METHOD PRIVATE Test_UnconnectedMon2IsRefused
TcUnit.TEST(__POUNAME());
// arrange / act: Mon2 is unconnected, which the Safety Editor refuses
group_3(Run := TRUE);
fb_3(Mon1 := TRUE);
group_3(Run := TRUE);
fb_3(Mon1 := TRUE);
// assert
AssertEquals_BOOL(Expected := TRUE, Actual := fb_3.Error, Message := 'configuration error reported');
AssertEquals_BYTE(Expected := TO_BYTE(E_SafeFbState.Error), Actual := fb_3.State, Message := 'state ERROR');
AssertEquals_WORD(Expected := WORD#16#8000, Actual := fb_3.Diag, Message := 'diag bit 15 configuration refused');
AssertEquals_BOOL(Expected := TRUE, Actual := group_3.FbErr, Message := 'the group sees an FB error');
// act: ErrAck 0 -> 1 -> 0 does not clear a configuration error
group_3(Run := TRUE, ErrAck := TRUE);
fb_3(Mon1 := TRUE);
group_3(Run := TRUE, ErrAck := TRUE);
fb_3(Mon1 := TRUE);
group_3(Run := TRUE, ErrAck := FALSE);
fb_3(Mon1 := TRUE);
AssertEquals_BOOL(Expected := TRUE, Actual := fb_3.Error, Message := 'error not acknowledged');
AssertEquals_WORD(Expected := WORD#16#8000, Actual := fb_3.Diag, Message := 'diag bit 15 kept');
TEST_FINISHED_NAMED(__POUNAME());
END_METHOD

END_FUNCTION_BLOCK

// ---- FunctionBlocks/T_SafeEdm.TcPOU
// Model of the TwinSAFE FB EDM (external device monitor):
// Mon2 must take the opposite value to Mon1 within the configured switch-on / switch-off time.
// The Safety Editor refuses an EDM with Mon1 or Mon2 unconnected: the model then reports Error with
// diagnostic bit 15 instead of running (see T_SafeFunctionBlockBase).
{attribute 'reflection'}
FUNCTION_BLOCK T_SafeEdm EXTENDS T_SafeFunctionBlockBase
VAR_INPUT
    Mon1 : BOOL;
    Mon2 : BOOL;
    Parameters : ST_SafeEdmParameters;
END_VAR
VAR
    {attribute 'is_connected' := 'Mon1'}
    _mon1Connected : BOOL;
    {attribute 'is_connected' := 'Mon2'}
    _mon2Connected : BOOL;
    _state : E_SafeEdmState := E_SafeEdmState.Stop;
    _prevState : E_SafeEdmState;
    _timer : TON;
    _satisfied : BOOL;
END_VAR

SUPER^();
IsRunning := (_state = E_SafeEdmState.MonOn) OR (_state = E_SafeEdmState.MonOff);

// Mon1 and Mon2 must both be connected (Safety Editor: "Inport Mon1 of EDM must be connected").
METHOD PROTECTED ConfigurationOk : BOOL
IF NOT _mon1Connected THEN
    _configurationFault := 'T_SafeEdm: Inport Mon1 of EDM must be connected';
    RETURN;
ELSIF NOT _mon2Connected THEN
    _configurationFault := 'T_SafeEdm: Inport Mon2 of EDM must be connected';
    RETURN;
END_IF

ConfigurationOk := TRUE;
END_METHOD

METHOD PROTECTED Process
VAR
    monitor1 : BOOL;
    monitor2 : BOOL;
    stateBefore : E_SafeEdmState;
    passes : USINT;
END_VAR
monitor1 := F_SafeInputValue(_mon1Connected, Parameters.Mon1MakeContact, Mon1);
monitor2 := F_SafeInputValue(_mon2Connected, Parameters.Mon2MakeContact, Mon2);

IF NOT _fbRun AND _state <> E_SafeEdmState.Error AND _state <> E_SafeEdmState.Reset THEN
    _state := E_SafeEdmState.Stop;
END_IF

passes := 0;

REPEAT
    stateBefore := _state;

    CASE _state OF
        E_SafeEdmState.Stop:
            IF StateChanged() THEN
                Error := FALSE;
                Diag  := 0;
                _timer(IN := FALSE, PT := T#0S);
            END_IF

            IF _fbRun THEN
                _state := SEL(monitor1, E_SafeEdmState.MonOff, E_SafeEdmState.MonOn);
            END_IF

        E_SafeEdmState.MonOn:
            // switch-on monitoring: Mon2 must become FALSE within SwitchOnTime
            IF StateChanged() THEN
                _satisfied := FALSE;
                _timer(IN := FALSE, PT := Parameters.SwitchOnTime);
            END_IF

            IF NOT monitor2 THEN
                _satisfied := TRUE;
            END_IF

            _timer(IN := NOT _satisfied AND (Parameters.SwitchOnTime > T#0S), PT := Parameters.SwitchOnTime);

            IF _timer.Q THEN
                SetDiagBit(1);
                _state := E_SafeEdmState.Error;
            ELSIF NOT monitor1 THEN
                _state := E_SafeEdmState.MonOff;
            END_IF

        E_SafeEdmState.MonOff:
            // switch-off monitoring: Mon2 must become TRUE within SwitchOffTime
            IF StateChanged() THEN
                _satisfied := FALSE;
                _timer(IN := FALSE, PT := Parameters.SwitchOffTime);
            END_IF

            IF monitor2 THEN
                _satisfied := TRUE;
            END_IF

            _timer(IN := NOT _satisfied AND (Parameters.SwitchOffTime > T#0S), PT := Parameters.SwitchOffTime);

            IF _timer.Q THEN
                SetDiagBit(0);
                _state := E_SafeEdmState.Error;
            ELSIF monitor1 THEN
                _state := E_SafeEdmState.MonOn;
            END_IF

        E_SafeEdmState.Error:
            IF StateChanged() THEN
                Error := TRUE;
                _timer(IN := FALSE, PT := T#0S);
            END_IF

            IF _errAck THEN
                _state := E_SafeEdmState.Reset;
            END_IF

        E_SafeEdmState.Reset:
            IF StateChanged() THEN
                Error := FALSE;
                Diag  := 0;
            END_IF

            IF _errAckFallingEdge THEN
                IF NOT _fbRun THEN
                    _state := E_SafeEdmState.Stop;
                ELSE
                    _state := SEL(monitor1, E_SafeEdmState.MonOff, E_SafeEdmState.MonOn);
                END_IF
            END_IF
    END_CASE

    passes := passes + 1;
UNTIL (stateBefore = _state) OR (passes >= 3)
END_REPEAT

State := TO_BYTE(_state);
END_METHOD

METHOD PRIVATE StateChanged : BOOL
IF _prevState = _state THEN
    RETURN;
END_IF

_prevState   := _state;
StateChanged := TRUE;
END_METHOD

END_FUNCTION_BLOCK

// ---- Tests/T_SafeEStop_Tests.TcPOU
FUNCTION_BLOCK T_SafeEStop_Tests EXTENDS TcUnit.FB_TestSuite
VAR
    // Test_OutputsOffWhenStopped
    group_1 : T_SafeGroup;
    fb_1 : T_SafeEStop(group := group_1);
    // Test_StartupRequiresRestartSequence
    group_2 : T_SafeGroup;
    fb_2 : T_SafeEStop(group := group_2);
    // Test_EStopRequestSwitchesOutputsOffAndBlocksRestart
    group_3 : T_SafeGroup;
    fb_3 : T_SafeEStop(group := group_3);
    // Test_MakeContactInputRequestsSafeStateOnOne
    group_4 : T_SafeGroup;
    fb_4 : T_SafeEStop(group := group_4) := (Parameters := (EStopIn1MakeContact := TRUE));
    // Test_EdmErrorAtRestartAndAcknowledge
    group_5 : T_SafeGroup;
    fb_5 : T_SafeEStop(group := group_5);
    // Test_RestartHeldBeforeEStopGivesEdmError
    group_6 : T_SafeGroup;
    fb_6 : T_SafeEStop(group := group_6);
    // Test_DelayedOutput
    group_7 : T_SafeGroup;
    fb_7 : T_SafeEStop(group := group_7) := (Parameters := (DelayTime := T#150MS));
    state_7 : INT := 10;
    waitTimer_7 : TON;
    // Test_DiscrepancyErrorNeedsSafeInputsBeforeAck
    group_8 : T_SafeGroup;
    fb_8 : T_SafeEStop(group := group_8) := (Parameters := (DiscrepancyTime1 := T#100MS));
    state_8 : INT := 10;
    waitTimer_8 : TON;
    // Test_ResetTimeOverSixtySecondsIsRefused
    group_9 : T_SafeGroup;
    fb_9 : T_SafeEStop(group := group_9) := (Parameters := (Edm2ResetTime := T#60010MS));
END_VAR

Test_OutputsOffWhenStopped();
Test_StartupRequiresRestartSequence();
Test_EStopRequestSwitchesOutputsOffAndBlocksRestart();
Test_MakeContactInputRequestsSafeStateOnOne();
Test_EdmErrorAtRestartAndAcknowledge();
Test_RestartHeldBeforeEStopGivesEdmError();
Test_DelayedOutput();
Test_DiscrepancyErrorNeedsSafeInputsBeforeAck();
Test_ResetTimeOverSixtySecondsIsRefused();

METHOD PRIVATE Test_DelayedOutput
TcUnit.TEST(__POUNAME());
waitTimer_7();

CASE state_7 OF
    10:
        // arrange: running
        group_7(Run := TRUE);
        fb_7(Restart := FALSE, EStopIn1 := TRUE);
        group_7(Run := TRUE);
        fb_7(Restart := TRUE, EStopIn1 := TRUE);
        group_7(Run := TRUE);
        fb_7(Restart := FALSE, EStopIn1 := TRUE);
        // act
        group_7(Run := TRUE);
        fb_7(Restart := FALSE, EStopIn1 := FALSE);
        // assert
        AssertEquals_BOOL(Expected := FALSE, Actual := fb_7.EStopOut, Message := 'EStopOut off immediately');
        AssertEquals_BOOL(Expected := TRUE, Actual := fb_7.EStopDelOut, Message := 'EStopDelOut still on');
        AssertEquals_BYTE(Expected := TO_BYTE(E_SafeFbState.DelayOut), Actual := fb_7.State, Message := 'state DELAYOUT');
        state_7 := 20;
        waitTimer_7(IN := TRUE, PT := T#300MS);
    20:
        group_7(Run := TRUE);
        fb_7(Restart := FALSE, EStopIn1 := FALSE);

        IF NOT waitTimer_7.Q THEN
            RETURN;
        END_IF

        waitTimer_7(IN := FALSE);
        // assert
        AssertEquals_BOOL(Expected := FALSE, Actual := fb_7.EStopDelOut, Message := 'EStopDelOut off after the delay');
        AssertEquals_BYTE(Expected := TO_BYTE(E_SafeFbState.Safe), Actual := fb_7.State, Message := 'state SAFE');
        TEST_FINISHED_NAMED(__POUNAME());
        state_7 := 10;
END_CASE
END_METHOD

METHOD PRIVATE Test_DiscrepancyErrorNeedsSafeInputsBeforeAck
TcUnit.TEST(__POUNAME());
waitTimer_8();

CASE state_8 OF
    10:
        // arrange: running
        group_8(Run := TRUE, ErrAck := FALSE);
        fb_8(Restart := FALSE, EStopIn1 := TRUE, EStopIn2 := TRUE);
        group_8(Run := TRUE, ErrAck := FALSE);
        fb_8(Restart := TRUE, EStopIn1 := TRUE, EStopIn2 := TRUE);
        group_8(Run := TRUE, ErrAck := FALSE);
        fb_8(Restart := FALSE, EStopIn1 := TRUE, EStopIn2 := TRUE);
        state_8 := 20;
        waitTimer_8(IN := TRUE, PT := T#250MS);
    20:
        // act: only one channel opens
        group_8(Run := TRUE, ErrAck := FALSE);
        fb_8(Restart := FALSE, EStopIn1 := FALSE, EStopIn2 := TRUE);

        IF NOT waitTimer_8.Q THEN
            RETURN;
        END_IF

        waitTimer_8(IN := FALSE);
        // assert
        AssertEquals_BOOL(Expected := TRUE, Actual := fb_8.Error, Message := 'discrepancy error');
        AssertEquals_WORD(Expected := WORD#16#0101, Actual := fb_8.Diag, Message := 'diag bits 0 and 8');
        // act: acknowledge while channel 2 is still closed
        group_8(Run := TRUE, ErrAck := TRUE);
        fb_8(Restart := FALSE, EStopIn1 := FALSE, EStopIn2 := TRUE);
        AssertEquals_BYTE(Expected := TO_BYTE(E_SafeFbState.Error), Actual := fb_8.State, Message := 'ack refused until both channels safe');
        group_8(Run := TRUE, ErrAck := TRUE);
        fb_8(Restart := FALSE, EStopIn1 := FALSE, EStopIn2 := FALSE);
        AssertEquals_BYTE(Expected := TO_BYTE(E_SafeFbState.Reset), Actual := fb_8.State, Message := 'RESET once both channels were safe');
        TEST_FINISHED_NAMED(__POUNAME());
        state_8 := 10;
END_CASE
END_METHOD

METHOD PRIVATE Test_EdmErrorAtRestartAndAcknowledge
TcUnit.TEST(__POUNAME());
// arrange: EDM1 connected but contactor not released
group_5(Run := TRUE, ErrAck := FALSE);
fb_5(Restart := FALSE, EDM1 := FALSE, EStopIn1 := TRUE);
// act: restart
group_5(Run := TRUE, ErrAck := FALSE);
fb_5(Restart := TRUE, EDM1 := FALSE, EStopIn1 := TRUE);
// assert
AssertEquals_BOOL(Expected := TRUE, Actual := fb_5.Error, Message := 'EDM error when feedback missing at restart');
AssertEquals_BYTE(Expected := TO_BYTE(E_SafeFbState.Error), Actual := fb_5.State, Message := 'state ERROR');
AssertEquals_WORD(Expected := WORD#16, Actual := fb_5.Diag, Message := 'diag bit 4 EDM1');
// act: the group_5 sees the error and leaves RUN; the FB error is held
group_5(Run := TRUE, ErrAck := FALSE);
fb_5(Restart := FALSE, EDM1 := FALSE, EStopIn1 := TRUE);
AssertEquals_BYTE(Expected := TO_BYTE(E_SafeGroupState.Error), Actual := group_5.State, Message := 'group ERROR');
AssertEquals_BYTE(Expected := TO_BYTE(E_SafeFbState.Error), Actual := fb_5.State, Message := 'error is held while the group is in ERROR');
// act: ErrAck 0 -> 1 (two cycles, the group_5 needs the second to reach RESET) -> 0
group_5(Run := TRUE, ErrAck := TRUE);
fb_5(Restart := FALSE, EDM1 := FALSE, EStopIn1 := TRUE);
AssertEquals_BYTE(Expected := TO_BYTE(E_SafeFbState.Reset), Actual := fb_5.State, Message := 'state RESET while ErrAck is 1');
AssertEquals_BOOL(Expected := FALSE, Actual := fb_5.Error, Message := 'Error output off in RESET');
group_5(Run := TRUE, ErrAck := TRUE);
fb_5(Restart := FALSE, EDM1 := FALSE, EStopIn1 := TRUE);
AssertEquals_BYTE(Expected := TO_BYTE(E_SafeGroupState.Reset), Actual := group_5.State, Message := 'group RESET');
group_5(Run := TRUE, ErrAck := FALSE);
fb_5(Restart := FALSE, EDM1 := FALSE, EStopIn1 := TRUE);
AssertEquals_BYTE(Expected := TO_BYTE(E_SafeGroupState.Run), Actual := group_5.State, Message := 'group RUN after ErrAck falling edge');
AssertEquals_BYTE(Expected := TO_BYTE(E_SafeFbState.Safe), Actual := fb_5.State, Message := 'state SAFE after ErrAck falling edge');
TEST_FINISHED_NAMED(__POUNAME());
END_METHOD

METHOD PRIVATE Test_EStopRequestSwitchesOutputsOffAndBlocksRestart
TcUnit.TEST(__POUNAME());
// arrange: running
group_3(Run := TRUE);
fb_3(Restart := FALSE, EStopIn1 := TRUE, EStopIn2 := TRUE);
group_3(Run := TRUE);
fb_3(Restart := TRUE, EStopIn1 := TRUE, EStopIn2 := TRUE);
group_3(Run := TRUE);
fb_3(Restart := FALSE, EStopIn1 := TRUE, EStopIn2 := TRUE);
// act: press the e-stop
group_3(Run := TRUE);
fb_3(Restart := FALSE, EStopIn1 := FALSE, EStopIn2 := FALSE);
// assert
AssertEquals_BOOL(Expected := FALSE, Actual := fb_3.EStopOut, Message := 'EStopOut off');
AssertEquals_BOOL(Expected := FALSE, Actual := fb_3.EStopDelOut, Message := 'EStopDelOut off without delay time');
AssertEquals_BYTE(Expected := TO_BYTE(E_SafeFbState.Safe), Actual := fb_3.State, Message := 'state SAFE');
// act: restart while still pressed
group_3(Run := TRUE);
fb_3(Restart := TRUE, EStopIn1 := FALSE, EStopIn2 := FALSE);
group_3(Run := TRUE);
fb_3(Restart := FALSE, EStopIn1 := FALSE, EStopIn2 := FALSE);
AssertEquals_BOOL(Expected := FALSE, Actual := fb_3.EStopOut, Message := 'restart ignored while the e-stop is pressed');
TEST_FINISHED_NAMED(__POUNAME());
END_METHOD

METHOD PRIVATE Test_MakeContactInputRequestsSafeStateOnOne
TcUnit.TEST(__POUNAME());
// arrange: single channel make contact, released (0), restarted
group_4(Run := TRUE);
fb_4(Restart := FALSE, EStopIn1 := FALSE);
group_4(Run := TRUE);
fb_4(Restart := TRUE, EStopIn1 := FALSE);
group_4(Run := TRUE);
fb_4(Restart := FALSE, EStopIn1 := FALSE);
AssertEquals_BYTE(Expected := TO_BYTE(E_SafeFbState.Run), Actual := fb_4.State, Message := 'running with make contact released');
// act
group_4(Run := TRUE);
fb_4(Restart := FALSE, EStopIn1 := TRUE);
// assert
AssertEquals_BYTE(Expected := TO_BYTE(E_SafeFbState.Safe), Actual := fb_4.State, Message := 'make contact at 1 requests the safe state');
TEST_FINISHED_NAMED(__POUNAME());
END_METHOD

METHOD PRIVATE Test_OutputsOffWhenStopped
TcUnit.TEST(__POUNAME());
// act
group_1(Run := FALSE);
fb_1(EStopIn1 := TRUE);
// assert
AssertEquals_BOOL(Expected := FALSE, Actual := fb_1.EStopOut, Message := 'no output while the group is stopped');
AssertEquals_BYTE(Expected := TO_BYTE(E_SafeFbState.Stop), Actual := fb_1.State, Message := 'state STOP');
TEST_FINISHED_NAMED(__POUNAME());
END_METHOD

METHOD PRIVATE Test_RestartHeldBeforeEStopGivesEdmError
TcUnit.TEST(__POUNAME());
// arrange: running with EDM feedback (contactors pulled in -> EDM1 = 0)
group_6(Run := TRUE);
fb_6(Restart := FALSE, EDM1 := TRUE, EStopIn1 := TRUE);
group_6(Run := TRUE);
fb_6(Restart := TRUE, EDM1 := TRUE, EStopIn1 := TRUE);
group_6(Run := TRUE);
fb_6(Restart := FALSE, EDM1 := TRUE, EStopIn1 := TRUE);
group_6(Run := TRUE);
fb_6(Restart := FALSE, EDM1 := FALSE, EStopIn1 := TRUE);
// act: restart held, then e-stop pressed before the contactors drop out
group_6(Run := TRUE);
fb_6(Restart := TRUE, EDM1 := FALSE, EStopIn1 := FALSE);
// assert
AssertEquals_BOOL(Expected := TRUE, Actual := fb_6.Error, Message := 'immediate EDM check with restart held (sample 3)');
TEST_FINISHED_NAMED(__POUNAME());
END_METHOD

METHOD PRIVATE Test_StartupRequiresRestartSequence
TcUnit.TEST(__POUNAME());
// act: two channel e-stop released, no restart yet
group_2(Run := TRUE);
fb_2(Restart := FALSE, EStopIn1 := TRUE, EStopIn2 := TRUE);
group_2(Run := TRUE);
fb_2(Restart := FALSE, EStopIn1 := TRUE, EStopIn2 := TRUE);
// assert
AssertEquals_BOOL(Expected := FALSE, Actual := fb_2.EStopOut, Message := 'no output before restart');
AssertEquals_BYTE(Expected := TO_BYTE(E_SafeFbState.Safe), Actual := fb_2.State, Message := 'state SAFE waiting for restart');
group_2(Run := TRUE);
fb_2(Restart := TRUE, EStopIn1 := TRUE, EStopIn2 := TRUE);
AssertEquals_BYTE(Expected := TO_BYTE(E_SafeFbState.Start), Actual := fb_2.State, Message := 'state START while restart held');
AssertEquals_BOOL(Expected := FALSE, Actual := fb_2.EStopOut, Message := 'no output while restart held');
group_2(Run := TRUE);
fb_2(Restart := FALSE, EStopIn1 := TRUE, EStopIn2 := TRUE);
AssertEquals_BYTE(Expected := TO_BYTE(E_SafeFbState.Run), Actual := fb_2.State, Message := 'state RUN after falling edge');
AssertEquals_BOOL(Expected := TRUE, Actual := fb_2.EStopOut, Message := 'EStopOut on');
AssertEquals_BOOL(Expected := TRUE, Actual := fb_2.EStopDelOut, Message := 'EStopDelOut on');
TEST_FINISHED_NAMED(__POUNAME());
END_METHOD

METHOD PRIVATE Test_ResetTimeOverSixtySecondsIsRefused
TcUnit.TEST(__POUNAME());
// arrange / act: Edm2ResetTime is 60010 ms, which the Safety Editor refuses
group_9(Run := TRUE);
fb_9(EDM2 := TRUE, EStopIn1 := TRUE);
group_9(Run := TRUE);
fb_9(EDM2 := TRUE, EStopIn1 := TRUE);
// assert
AssertEquals_BOOL(Expected := TRUE, Actual := fb_9.Error, Message := 'configuration error reported');
AssertEquals_BYTE(Expected := TO_BYTE(E_SafeFbState.Error), Actual := fb_9.State, Message := 'state ERROR');
AssertEquals_WORD(Expected := WORD#16#8000, Actual := fb_9.Diag, Message := 'diag bit 15 configuration refused');
AssertEquals_BOOL(Expected := FALSE, Actual := fb_9.EStopOut, Message := 'EStopOut stays at its safe value');
AssertEquals_BOOL(Expected := TRUE, Actual := group_9.FbErr, Message := 'the group sees an FB error');
// act: ErrAck 0 -> 1 -> 0 does not clear a configuration error
group_9(Run := TRUE, ErrAck := TRUE);
fb_9(EDM2 := TRUE, EStopIn1 := TRUE);
group_9(Run := TRUE, ErrAck := TRUE);
fb_9(EDM2 := TRUE, EStopIn1 := TRUE);
group_9(Run := TRUE, ErrAck := FALSE);
fb_9(EDM2 := TRUE, EStopIn1 := TRUE);
AssertEquals_BOOL(Expected := TRUE, Actual := fb_9.Error, Message := 'error not acknowledged');
AssertEquals_WORD(Expected := WORD#16#8000, Actual := fb_9.Diag, Message := 'diag bit 15 kept');
TEST_FINISHED_NAMED(__POUNAME());
END_METHOD

END_FUNCTION_BLOCK

// ---- FunctionBlocks/T_SafeEStop.TcPOU
// Model of the TwinSAFE FB ESTOP.
// Up to eight emergency stop inputs in four pairs, immediate and delayed outputs,
// two feedback loops (EDM) and a manual restart requiring a 0 -> 1 -> 0 sequence on Restart.
// Ports are active when connected.
// The Safety Editor refuses an EDM reset time that is not 0 ms, a multiple of 10 ms and at most 60000 ms:
// the model then reports Error with diagnostic bit 15 instead of running (see T_SafeFunctionBlockBase).
{attribute 'reflection'}
FUNCTION_BLOCK T_SafeEStop EXTENDS T_SafeFunctionBlockBase
VAR_INPUT
    Restart : BOOL; // may be a standard PLC signal
    EDM1 : BOOL; // feedback loop of EStopOut (may be a standard PLC signal)
    EDM2 : BOOL; // feedback loop of EStopDelOut (may be a standard PLC signal)
    EStopIn1 : BOOL;
    EStopIn2 : BOOL;
    EStopIn3 : BOOL;
    EStopIn4 : BOOL;
    EStopIn5 : BOOL;
    EStopIn6 : BOOL;
    EStopIn7 : BOOL;
    EStopIn8 : BOOL;
    Parameters : ST_SafeEStopParameters;
END_VAR
VAR_OUTPUT
    EStopOut : BOOL; // switches off immediately
    EStopDelOut : BOOL; // switches off after DelayTime
END_VAR
VAR
    {attribute 'is_connected' := 'Restart'}
    _restartConnected : BOOL;
    {attribute 'is_connected' := 'EDM1'}
    _eDM1Connected : BOOL;
    {attribute 'is_connected' := 'EDM2'}
    _eDM2Connected : BOOL;
    {attribute 'is_connected' := 'EStopIn1'}
    _eStopIn1Connected : BOOL;
    {attribute 'is_connected' := 'EStopIn2'}
    _eStopIn2Connected : BOOL;
    {attribute 'is_connected' := 'EStopIn3'}
    _eStopIn3Connected : BOOL;
    {attribute 'is_connected' := 'EStopIn4'}
    _eStopIn4Connected : BOOL;
    {attribute 'is_connected' := 'EStopIn5'}
    _eStopIn5Connected : BOOL;
    {attribute 'is_connected' := 'EStopIn6'}
    _eStopIn6Connected : BOOL;
    {attribute 'is_connected' := 'EStopIn7'}
    _eStopIn7Connected : BOOL;
    {attribute 'is_connected' := 'EStopIn8'}
    _eStopIn8Connected : BOOL;
    _pairs : ARRAY[1..4] OF T_SafeInputPair;
    _state : E_SafeFbState := E_SafeFbState.Stop;
    _prevState : E_SafeFbState;
    _restartPrev : BOOL;
    _delayTimer : TON;
    _edmResetTimer1 : TON;
    _edmResetTimer2 : TON;
    _edm1Dropped : BOOL;
    _edm2Dropped : BOOL;
END_VAR

SUPER^();

// The EDM reset times must be 0 ms or a multiple of 10 ms up to 60000 ms (Safety Editor: "'Reset Time' parameter ... has to be 0 ms or a multiple of 10 ms and maximal 60000 ms").
METHOD PROTECTED ConfigurationOk : BOOL
IF NOT F_SafeResetTimeOk(Parameters.Edm1ResetTime) THEN
    _configurationFault := 'T_SafeEStop: $'Reset Time$' parameter of EDM1 of ESTOP has to be 0 ms or a multiple of 10 ms and maximal 60000 ms';
    RETURN;
ELSIF NOT F_SafeResetTimeOk(Parameters.Edm2ResetTime) THEN
    _configurationFault := 'T_SafeEStop: $'Reset Time$' parameter of EDM2 of ESTOP has to be 0 ms or a multiple of 10 ms and maximal 60000 ms';
    RETURN;
END_IF

ConfigurationOk := TRUE;
END_METHOD

// Checks the EDM inputs at restart and records diagnostic bits 4/5 on failure.
METHOD PRIVATE EdmInputsOk : BOOL
EdmInputsOk := TRUE;

IF _eDM1Connected AND NOT EDM1 THEN
    SetDiagBit(4);
    EdmInputsOk := FALSE;
END_IF

IF _eDM2Connected AND NOT EDM2 THEN
    SetDiagBit(5);
    EdmInputsOk := FALSE;
END_IF
END_METHOD

// TRUE when every connected EDM input reads 1 (contactors released).
METHOD PRIVATE EdmInputsTrue : BOOL
EdmInputsTrue := (NOT _eDM1Connected OR EDM1) AND (NOT _eDM2Connected OR EDM2);
END_METHOD

// EL6910 extension: after the outputs switch on, each connected EDM input must drop to FALSE
// within its Reset Time. Returns FALSE (and sets diagnostic bits 4/5) on timeout.
METHOD PRIVATE EdmResetOk : BOOL
EdmResetOk := TRUE;

IF _eDM1Connected AND Parameters.Edm1ResetTime > T#0S THEN
    IF NOT EDM1 THEN
        _edm1Dropped := TRUE;
    END_IF

    _edmResetTimer1(IN := NOT _edm1Dropped, PT := Parameters.Edm1ResetTime);

    IF _edmResetTimer1.Q THEN
        SetDiagBit(4);
        EdmResetOk := FALSE;
    END_IF
END_IF

IF _eDM2Connected AND Parameters.Edm2ResetTime > T#0S THEN
    IF NOT EDM2 THEN
        _edm2Dropped := TRUE;
    END_IF

    _edmResetTimer2(IN := NOT _edm2Dropped, PT := Parameters.Edm2ResetTime);

    IF _edmResetTimer2.Q THEN
        SetDiagBit(5);
        EdmResetOk := FALSE;
    END_IF
END_IF
END_METHOD

PROPERTY EStopState : E_SafeFbState
GET
EStopState := _state;
END_GET
END_PROPERTY

METHOD PROTECTED Process
VAR
    i : USINT;
    acknowledge : BOOL;
    safeRequested : BOOL;
    discError : BOOL;
    restartFalling : BOOL;
    operating : BOOL;
    stateBefore : E_SafeFbState;
    passes : USINT;
END_VAR
acknowledge := (_state = E_SafeFbState.Error) AND _errAck;
_pairs[1](
    In1 := EStopIn1,
    In2 := EStopIn2,
    Active1 := _eStopIn1Connected,
    Active2 := _eStopIn2Connected,
    MakeContact1 := Parameters.EStopIn1MakeContact,
    MakeContact2 := Parameters.EStopIn2MakeContact,
    DiscrepancyTime := Parameters.DiscrepancyTime1,
    Monitor := _fbRun,
    SafeInputsAfterDiscError := TRUE, // the EL6910 always applies it to ESTOP, whatever the parameter says
    Acknowledge := acknowledge
);

_pairs[2](
    In1 := EStopIn3,
    In2 := EStopIn4,
    Active1 := _eStopIn3Connected,
    Active2 := _eStopIn4Connected,
    MakeContact1 := Parameters.EStopIn3MakeContact,
    MakeContact2 := Parameters.EStopIn4MakeContact,
    DiscrepancyTime := Parameters.DiscrepancyTime2,
    Monitor := _fbRun,
    SafeInputsAfterDiscError := TRUE, // the EL6910 always applies it to ESTOP, whatever the parameter says
    Acknowledge := acknowledge
);

_pairs[3](
    In1 := EStopIn5,
    In2 := EStopIn6,
    Active1 := _eStopIn5Connected,
    Active2 := _eStopIn6Connected,
    MakeContact1 := Parameters.EStopIn5MakeContact,
    MakeContact2 := Parameters.EStopIn6MakeContact,
    DiscrepancyTime := Parameters.DiscrepancyTime3,
    Monitor := _fbRun,
    SafeInputsAfterDiscError := TRUE, // the EL6910 always applies it to ESTOP, whatever the parameter says
    Acknowledge := acknowledge
);

_pairs[4](
    In1 := EStopIn7,
    In2 := EStopIn8,
    Active1 := _eStopIn7Connected,
    Active2 := _eStopIn8Connected,
    MakeContact1 := Parameters.EStopIn7MakeContact,
    MakeContact2 := Parameters.EStopIn8MakeContact,
    DiscrepancyTime := Parameters.DiscrepancyTime4,
    Monitor := _fbRun,
    SafeInputsAfterDiscError := TRUE, // the EL6910 always applies it to ESTOP, whatever the parameter says
    Acknowledge := acknowledge
);

FOR i := 1 TO 4 DO
    safeRequested := safeRequested OR _pairs[i].SafeStateRequested;
    discError     := discError OR _pairs[i].DiscrepancyError;
END_FOR

restartFalling := NOT Restart AND _restartPrev;
_restartPrev   := Restart;

IF NOT _fbRun AND _state <> E_SafeFbState.Error AND _state <> E_SafeFbState.Reset THEN
    _state := E_SafeFbState.Stop;
END_IF

// A discrepancy error is detected in every operating state
operating := (_state = E_SafeFbState.Safe)
                 OR (_state = E_SafeFbState.Start)
                 OR (_state = E_SafeFbState.Run)
                 OR (_state = E_SafeFbState.DelayOut);

IF discError AND operating THEN
    UpdateDiscrepancyDiag();
    _state := E_SafeFbState.Error;
END_IF

passes := 0;

REPEAT
    stateBefore := _state;

    CASE _state OF
        E_SafeFbState.Stop:
            IF StateChanged() THEN
                SetOutputsSafe();
                Error := FALSE;
                Diag  := 0;
            END_IF

            IF _fbRun THEN
                _state := E_SafeFbState.Safe;
            END_IF

        E_SafeFbState.Safe:
            IF StateChanged() THEN
                SetOutputsSafe();
            END_IF

            // A TRUE restart signal triggers the EDM check immediately (see restart behaviour sample 3)
            IF Restart THEN
                IF NOT EdmInputsOk() THEN
                    _state := E_SafeFbState.Error;
                ELSIF NOT safeRequested THEN
                    _state := E_SafeFbState.Start;
                END_IF
            END_IF

        E_SafeFbState.Start:
            IF StateChanged() THEN
                SetOutputsSafe();
            END_IF

            IF safeRequested THEN
                _state := E_SafeFbState.Safe;
            ELSIF restartFalling THEN
                IF EdmInputsOk() THEN
                    _state := E_SafeFbState.Run;
                ELSE
                    _state := E_SafeFbState.Error;
                END_IF
            END_IF

        E_SafeFbState.Run:
            IF StateChanged() THEN
                EStopOut    := TRUE;
                EStopDelOut := TRUE;
                StartEdmResetMonitoring();
            END_IF

            IF NOT EdmResetOk() THEN
                _state := E_SafeFbState.Error;
            ELSIF safeRequested THEN
                IF Parameters.DelayTime > T#0S THEN
                    _state := E_SafeFbState.DelayOut;
                ELSE
                    _state := E_SafeFbState.Safe;
                END_IF
            END_IF

        E_SafeFbState.DelayOut:
            IF StateChanged() THEN
                EStopOut    := FALSE;
                EStopDelOut := TRUE;
                _delayTimer(IN := FALSE, PT := Parameters.DelayTime);
            END_IF

            _delayTimer(IN := TRUE, PT := Parameters.DelayTime);

            IF _delayTimer.Q THEN
                _state := E_SafeFbState.Safe;
            END_IF

        E_SafeFbState.Error:
            IF StateChanged() THEN
                SetOutputsSafe();
                Error := TRUE;
            END_IF

            UpdateDiscrepancyDiag();

            IF _errAck AND NOT discError THEN
                _state := E_SafeFbState.Reset;
            END_IF

        E_SafeFbState.Reset:
            IF StateChanged() THEN
                SetOutputsSafe();
                Error := FALSE;
                Diag  := 0;
            END_IF

            IF _errAckFallingEdge THEN
                _state := SEL(_fbRun, E_SafeFbState.Stop, E_SafeFbState.Safe);
            END_IF
    END_CASE

    passes := passes + 1;
UNTIL (stateBefore = _state) OR (passes >= 3)
END_REPEAT

State := TO_BYTE(_state);
END_METHOD

METHOD PRIVATE SetOutputsSafe
EStopOut    := FALSE;
EStopDelOut := FALSE;
END_METHOD

METHOD PRIVATE StartEdmResetMonitoring
_edm1Dropped := FALSE;
_edm2Dropped := FALSE;
_edmResetTimer1(IN := FALSE, PT := Parameters.Edm1ResetTime);
_edmResetTimer2(IN := FALSE, PT := Parameters.Edm2ResetTime);
END_METHOD

METHOD PRIVATE StateChanged : BOOL
IF _prevState = _state THEN
    RETURN;
END_IF

_prevState   := _state;
StateChanged := TRUE;
END_METHOD

// Mirrors the discrepancy state of every pair into the diagnostic bits.
METHOD PRIVATE UpdateDiscrepancyDiag
VAR
    i : USINT;
END_VAR
FOR i := 1 TO 4 DO
    IF _pairs[i].DiscrepancyError THEN
        SetDiagBit(i - 1);

        IF _pairs[i].AwaitingSafeInputs THEN
            SetDiagBit(i + 7);
        ELSE
            ClearDiagBit(i + 7);
        END_IF
    END_IF
END_FOR
END_METHOD

END_FUNCTION_BLOCK

// ---- Core/F_SafeResetTimeOk.TcPOU
// TRUE when an EDM 'Reset Time' parameter is one the Safety Editor accepts: 0 ms (off) or a multiple
// of 10 ms, and at most 60000 ms. The editor reports "'Reset Time' parameter ... has to be 0 ms or a
// multiple of 10 ms and maximal 60000 ms" otherwise.
FUNCTION F_SafeResetTimeOk : BOOL
VAR_INPUT
    resetTime : TIME;
END_VAR
VAR CONSTANT
    MAX_RESET_TIME : TIME := T#60S;
END_VAR

IF resetTime > MAX_RESET_TIME THEN
    RETURN;
END_IF

F_SafeResetTimeOk := (TIME_TO_UDINT(resetTime) MOD 10 = 0);

END_FUNCTION

// ---- Tests/T_SafeMon_Tests.TcPOU
FUNCTION_BLOCK T_SafeMon_Tests EXTENDS TcUnit.FB_TestSuite
VAR
    // Test_AutomaticRestartWhenGuardClosed
    group_1 : T_SafeGroup;
    fb_1 : T_SafeMon(group := group_1);
    // Test_SecureInputBypassesGuard
    group_2 : T_SafeGroup;
    fb_2 : T_SafeMon(group := group_2);
    // Test_ManualFunctionTestRequiresGuardOpenedOnce
    group_3 : T_SafeGroup;
    fb_3 : T_SafeMon(group := group_3) := (Parameters := (ManualFunctionTest := TRUE));
    // Test_EdmFaultWithoutManualRestartStaysSafe
    group_4 : T_SafeGroup;
    fb_4 : T_SafeMon(group := group_4);
    // Test_NoMonInConnectedIsRefused
    group_5 : T_SafeGroup;
    fb_5 : T_SafeMon(group := group_5);
    // Test_ResetTimeNotMultipleOfTenIsRefused
    group_6 : T_SafeGroup;
    fb_6 : T_SafeMon(group := group_6) := (Parameters := (Edm1ResetTime := T#15MS));
END_VAR

Test_AutomaticRestartWhenGuardClosed();
Test_SecureInputBypassesGuard();
Test_ManualFunctionTestRequiresGuardOpenedOnce();
Test_EdmFaultWithoutManualRestartStaysSafe();
Test_NoMonInConnectedIsRefused();
Test_ResetTimeNotMultipleOfTenIsRefused();

METHOD PRIVATE Test_AutomaticRestartWhenGuardClosed
TcUnit.TEST(__POUNAME());
// act: Restart not connected -> automatic restart; guard open
group_1(Run := TRUE);
fb_1(MonIn1 := FALSE);
group_1(Run := TRUE);
fb_1(MonIn1 := FALSE);
// assert
AssertEquals_BOOL(Expected := FALSE, Actual := fb_1.MonOut, Message := 'output off with guard open');
group_1(Run := TRUE);
fb_1(MonIn1 := TRUE);
AssertEquals_BOOL(Expected := TRUE, Actual := fb_1.MonOut, Message := 'automatic restart with guard closed');
AssertEquals_BYTE(Expected := TO_BYTE(E_SafeMonState.Run), Actual := fb_1.State, Message := 'state RUN');
TEST_FINISHED_NAMED(__POUNAME());
END_METHOD

METHOD PRIVATE Test_EdmFaultWithoutManualRestartStaysSafe
TcUnit.TEST(__POUNAME());
// act: EDM1 connected and FALSE, no Restart connected
group_4(Run := TRUE);
fb_4(EDM1 := FALSE, MonIn1 := TRUE);
group_4(Run := TRUE);
fb_4(EDM1 := FALSE, MonIn1 := TRUE);
// assert
AssertEquals_BOOL(Expected := FALSE, Actual := fb_4.Error, Message := 'no EDM error without manual restart');
AssertEquals_BYTE(Expected := TO_BYTE(E_SafeMonState.Safe), Actual := fb_4.State, Message := 'FB remains SAFE');
TEST_FINISHED_NAMED(__POUNAME());
END_METHOD

METHOD PRIVATE Test_ManualFunctionTestRequiresGuardOpenedOnce
TcUnit.TEST(__POUNAME());
// arrange: Restart connected (manual restart), guard closed from the start
group_3(Run := TRUE);
fb_3(Restart := FALSE, MonIn1 := TRUE);
AssertEquals_BYTE(Expected := TO_BYTE(E_SafeMonState.FuncTest), Actual := fb_3.State, Message := 'state FUNCTEST after start');
// act: restart without testing the guard
group_3(Run := TRUE);
fb_3(Restart := TRUE, MonIn1 := TRUE);
group_3(Run := TRUE);
fb_3(Restart := FALSE, MonIn1 := TRUE);
AssertEquals_BOOL(Expected := FALSE, Actual := fb_3.MonOut, Message := 'restart ignored before the function test');
// act: open and close the guard, then restart
group_3(Run := TRUE);
fb_3(Restart := FALSE, MonIn1 := FALSE);
group_3(Run := TRUE);
fb_3(Restart := FALSE, MonIn1 := TRUE);
group_3(Run := TRUE);
fb_3(Restart := TRUE, MonIn1 := TRUE);
group_3(Run := TRUE);
fb_3(Restart := FALSE, MonIn1 := TRUE);
AssertEquals_BOOL(Expected := TRUE, Actual := fb_3.MonOut, Message := 'output on after function test and restart');
TEST_FINISHED_NAMED(__POUNAME());
END_METHOD

METHOD PRIVATE Test_SecureInputBypassesGuard
TcUnit.TEST(__POUNAME());
// act: guard open, bypass active
group_2(Run := TRUE);
fb_2(MonIn1 := FALSE, Secure1 := TRUE);
group_2(Run := TRUE);
fb_2(MonIn1 := FALSE, Secure1 := TRUE);
// assert
AssertEquals_BOOL(Expected := TRUE, Actual := fb_2.MonOut, Message := 'guard ignored while Secure is 1');
group_2(Run := TRUE);
fb_2(MonIn1 := FALSE, Secure1 := FALSE);
AssertEquals_BOOL(Expected := FALSE, Actual := fb_2.MonOut, Message := 'guard monitored again when Secure is 0');
TEST_FINISHED_NAMED(__POUNAME());
END_METHOD

METHOD PRIVATE Test_NoMonInConnectedIsRefused
TcUnit.TEST(__POUNAME());
// arrange / act: only the Secure pair is connected, which the Safety Editor refuses
group_5(Run := TRUE);
fb_5(Secure1 := TRUE);
group_5(Run := TRUE);
fb_5(Secure1 := TRUE);
// assert
AssertEquals_BOOL(Expected := TRUE, Actual := fb_5.Error, Message := 'configuration error reported');
AssertEquals_BYTE(Expected := TO_BYTE(E_SafeFbState.Error), Actual := fb_5.State, Message := 'state ERROR');
AssertEquals_WORD(Expected := WORD#16#8000, Actual := fb_5.Diag, Message := 'diag bit 15 configuration refused');
AssertEquals_BOOL(Expected := FALSE, Actual := fb_5.MonOut, Message := 'MonOut stays at its safe value');
AssertEquals_BOOL(Expected := TRUE, Actual := group_5.FbErr, Message := 'the group sees an FB error');
// act: ErrAck 0 -> 1 -> 0 does not clear a configuration error
group_5(Run := TRUE, ErrAck := TRUE);
fb_5(Secure1 := TRUE);
group_5(Run := TRUE, ErrAck := TRUE);
fb_5(Secure1 := TRUE);
group_5(Run := TRUE, ErrAck := FALSE);
fb_5(Secure1 := TRUE);
AssertEquals_BOOL(Expected := TRUE, Actual := fb_5.Error, Message := 'error not acknowledged');
AssertEquals_WORD(Expected := WORD#16#8000, Actual := fb_5.Diag, Message := 'diag bit 15 kept');
TEST_FINISHED_NAMED(__POUNAME());
END_METHOD

METHOD PRIVATE Test_ResetTimeNotMultipleOfTenIsRefused
TcUnit.TEST(__POUNAME());
// arrange / act: Edm1ResetTime is 15 ms, which the Safety Editor refuses
group_6(Run := TRUE);
fb_6(EDM1 := TRUE, MonIn1 := TRUE);
group_6(Run := TRUE);
fb_6(EDM1 := TRUE, MonIn1 := TRUE);
// assert
AssertEquals_BOOL(Expected := TRUE, Actual := fb_6.Error, Message := 'configuration error reported');
AssertEquals_BYTE(Expected := TO_BYTE(E_SafeFbState.Error), Actual := fb_6.State, Message := 'state ERROR');
AssertEquals_WORD(Expected := WORD#16#8000, Actual := fb_6.Diag, Message := 'diag bit 15 configuration refused');
AssertEquals_BOOL(Expected := FALSE, Actual := fb_6.MonOut, Message := 'MonOut stays at its safe value');
AssertEquals_BOOL(Expected := TRUE, Actual := group_6.FbErr, Message := 'the group sees an FB error');
// act: ErrAck 0 -> 1 -> 0 does not clear a configuration error
group_6(Run := TRUE, ErrAck := TRUE);
fb_6(EDM1 := TRUE, MonIn1 := TRUE);
group_6(Run := TRUE, ErrAck := TRUE);
fb_6(EDM1 := TRUE, MonIn1 := TRUE);
group_6(Run := TRUE, ErrAck := FALSE);
fb_6(EDM1 := TRUE, MonIn1 := TRUE);
AssertEquals_BOOL(Expected := TRUE, Actual := fb_6.Error, Message := 'error not acknowledged');
AssertEquals_WORD(Expected := WORD#16#8000, Actual := fb_6.Diag, Message := 'diag bit 15 kept');
TEST_FINISHED_NAMED(__POUNAME());
END_METHOD

END_FUNCTION_BLOCK

// ---- FunctionBlocks/T_SafeMon.TcPOU
// Model of the TwinSAFE FB MON (safety door / guard monitoring).
// Two MonIn pairs, a Secure pair that bypasses them, manual restart (when Restart is connected),
// manual function test, two EDM feedback loops and a delayed output.
// The Safety Editor refuses a MON with no MonIn port connected, or an EDM reset time that is not 0 ms,
// a multiple of 10 ms and at most 60000 ms: the model then reports Error with diagnostic bit 15
// instead of running (see T_SafeFunctionBlockBase).
{attribute 'reflection'}
FUNCTION_BLOCK T_SafeMon EXTENDS T_SafeFunctionBlockBase
VAR_INPUT
    Restart : BOOL; // connect for manual restart; may be a standard PLC signal
    EDM1 : BOOL; // feedback loop of MonOut
    EDM2 : BOOL; // feedback loop of MonDelOut
    MonIn1 : BOOL;
    MonIn2 : BOOL;
    MonIn3 : BOOL;
    MonIn4 : BOOL;
    Secure1 : BOOL; // when TRUE (after normalisation) the MonIn inputs are ignored
    Secure2 : BOOL;
    Parameters : ST_SafeMonParameters;
END_VAR
VAR_OUTPUT
    MonOut : BOOL;
    MonDelOut : BOOL;
END_VAR
VAR
    {attribute 'is_connected' := 'Restart'}
    _restartConnected : BOOL;
    {attribute 'is_connected' := 'EDM1'}
    _eDM1Connected : BOOL;
    {attribute 'is_connected' := 'EDM2'}
    _eDM2Connected : BOOL;
    {attribute 'is_connected' := 'MonIn1'}
    _monIn1Connected : BOOL;
    {attribute 'is_connected' := 'MonIn2'}
    _monIn2Connected : BOOL;
    {attribute 'is_connected' := 'MonIn3'}
    _monIn3Connected : BOOL;
    {attribute 'is_connected' := 'MonIn4'}
    _monIn4Connected : BOOL;
    {attribute 'is_connected' := 'Secure1'}
    _secure1Connected : BOOL;
    {attribute 'is_connected' := 'Secure2'}
    _secure2Connected : BOOL;
    _pairs : ARRAY[1..3] OF T_SafeInputPair; // 1: MonIn1/2, 2: MonIn3/4, 3: Secure1/2
    _state : E_SafeMonState := E_SafeMonState.Stop;
    _prevState : E_SafeMonState;
    _restartPrev : BOOL;
    _delayTimer : TON;
    _delayRunning : BOOL;
    _funcTested : ARRAY[1..2] OF BOOL;
    _edmResetTimer1 : TON;
    _edmResetTimer2 : TON;
    _edm1Dropped : BOOL;
    _edm2Dropped : BOOL;
END_VAR

SUPER^();

// At least one MonIn port must be connected and the EDM reset times must be 0 ms or a multiple of 10 ms up to 60000 ms (Safety Editor messages).
METHOD PROTECTED ConfigurationOk : BOOL
IF NOT (_monIn1Connected OR _monIn2Connected OR _monIn3Connected OR _monIn4Connected) THEN
    _configurationFault := 'T_SafeMon: MON does not have at least 1 MonIn(x) port active and connected';
    RETURN;
ELSIF NOT F_SafeResetTimeOk(Parameters.Edm1ResetTime) THEN
    _configurationFault := 'T_SafeMon: $'Reset Time$' parameter of EDM1 of MON has to be 0 ms or a multiple of 10 ms and maximal 60000 ms';
    RETURN;
ELSIF NOT F_SafeResetTimeOk(Parameters.Edm2ResetTime) THEN
    _configurationFault := 'T_SafeMon: $'Reset Time$' parameter of EDM2 of MON has to be 0 ms or a multiple of 10 ms and maximal 60000 ms';
    RETURN;
END_IF

ConfigurationOk := TRUE;
END_METHOD

// Checks the EDM inputs at restart and records diagnostic bits 4/5 on failure.
METHOD PRIVATE EdmInputsOk : BOOL
EdmInputsOk := TRUE;

IF _eDM1Connected AND NOT EDM1 THEN
    SetDiagBit(4);
    EdmInputsOk := FALSE;
END_IF

IF _eDM2Connected AND NOT EDM2 THEN
    SetDiagBit(5);
    EdmInputsOk := FALSE;
END_IF
END_METHOD

// TRUE when every connected EDM input reads 1 (contactors released).
METHOD PRIVATE EdmInputsTrue : BOOL
EdmInputsTrue := (NOT _eDM1Connected OR EDM1) AND (NOT _eDM2Connected OR EDM2);
END_METHOD

// EL6910 extension: after the outputs switch on, each connected EDM input must drop to FALSE
// within its Reset Time. Returns FALSE (and sets diagnostic bits 4/5) on timeout.
METHOD PRIVATE EdmResetOk : BOOL
EdmResetOk := TRUE;

IF _eDM1Connected AND Parameters.Edm1ResetTime > T#0S THEN
    IF NOT EDM1 THEN
        _edm1Dropped := TRUE;
    END_IF

    _edmResetTimer1(IN := NOT _edm1Dropped, PT := Parameters.Edm1ResetTime);

    IF _edmResetTimer1.Q THEN
        SetDiagBit(4);
        EdmResetOk := FALSE;
    END_IF
END_IF

IF _eDM2Connected AND Parameters.Edm2ResetTime > T#0S THEN
    IF NOT EDM2 THEN
        _edm2Dropped := TRUE;
    END_IF

    _edmResetTimer2(IN := NOT _edm2Dropped, PT := Parameters.Edm2ResetTime);

    IF _edmResetTimer2.Q THEN
        SetDiagBit(5);
        EdmResetOk := FALSE;
    END_IF
END_IF
END_METHOD

PROPERTY MonState : E_SafeMonState
GET
MonState := _state;
END_GET
END_PROPERTY

METHOD PROTECTED Process
VAR
    i : USINT;
    acknowledge : BOOL;
    monRequested : BOOL;
    bypass : BOOL;
    safeRequested : BOOL;
    discError : BOOL;
    restartFalling : BOOL;
    functionTestDue : BOOL;
    stateBefore : E_SafeMonState;
    passes : USINT;
END_VAR
acknowledge := (_state = E_SafeMonState.Error) AND _errAck;
_pairs[1](
    In1 := MonIn1,
    In2 := MonIn2,
    Active1 := _monIn1Connected,
    Active2 := _monIn2Connected,
    MakeContact1 := Parameters.MonIn1MakeContact,
    MakeContact2 := Parameters.MonIn2MakeContact,
    DiscrepancyTime := Parameters.DiscrepancyTime1,
    Monitor := _fbRun,
    SafeInputsAfterDiscError := Parameters.SafeInputsAfterDiscError,
    Acknowledge := acknowledge
);

_pairs[2](
    In1 := MonIn3,
    In2 := MonIn4,
    Active1 := _monIn3Connected,
    Active2 := _monIn4Connected,
    MakeContact1 := Parameters.MonIn3MakeContact,
    MakeContact2 := Parameters.MonIn4MakeContact,
    DiscrepancyTime := Parameters.DiscrepancyTime2,
    Monitor := _fbRun,
    SafeInputsAfterDiscError := Parameters.SafeInputsAfterDiscError,
    Acknowledge := acknowledge
);

_pairs[3](
    In1 := Secure1,
    In2 := Secure2,
    Active1 := _secure1Connected,
    Active2 := _secure2Connected,
    MakeContact1 := Parameters.Secure1MakeContact,
    MakeContact2 := Parameters.Secure2MakeContact,
    DiscrepancyTime := Parameters.SecureDiscrepancyTime,
    Monitor := _fbRun,
    SafeInputsAfterDiscError := Parameters.SafeInputsAfterDiscError,
    Acknowledge := acknowledge
);

monRequested  := _pairs[1].SafeStateRequested OR _pairs[2].SafeStateRequested;
bypass        := _pairs[3].IsActive AND _pairs[3].AllTrue;
safeRequested := monRequested AND NOT bypass;

FOR i := 1 TO 3 DO
    discError := discError OR _pairs[i].DiscrepancyError;
END_FOR

restartFalling := NOT Restart AND _restartPrev;
_restartPrev   := Restart;

IF NOT _fbRun AND _state <> E_SafeMonState.Error AND _state <> E_SafeMonState.Reset THEN
    _state := E_SafeMonState.Stop;
END_IF

// Discrepancy errors: immediate, except that a running delayed output completes its delay first
IF discError THEN
    CASE _state OF
        E_SafeMonState.Safe, E_SafeMonState.Start, E_SafeMonState.FuncTest:
            UpdateDiscrepancyDiag();
            _state := E_SafeMonState.Error;
        E_SafeMonState.Run:
            UpdateDiscrepancyDiag();

            IF Parameters.DelayTime > T#0S THEN
                _state := E_SafeMonState.ErrorDelay;
            ELSE
                _state := E_SafeMonState.Error;
            END_IF
        E_SafeMonState.DelayOut:
            UpdateDiscrepancyDiag();
            _state := E_SafeMonState.ErrorDelay;
    END_CASE
END_IF

passes := 0;

REPEAT
    stateBefore := _state;

    CASE _state OF
        E_SafeMonState.Stop:
            IF StateChanged() THEN
                SetOutputsSafe();
                Error          := FALSE;
                Diag           := 0;
                _delayRunning  := FALSE;
                _funcTested[1] := FALSE;
                _funcTested[2] := FALSE;
            END_IF

            IF _fbRun THEN
                functionTestDue := Parameters.ManualFunctionTest AND (_pairs[1].IsActive OR _pairs[2].IsActive);
                _state          := SEL(functionTestDue, E_SafeMonState.Safe, E_SafeMonState.FuncTest);
            END_IF

        E_SafeMonState.FuncTest:
            // every connected MonIn pair must request the safe state once before a restart is accepted
            IF StateChanged() THEN
                SetOutputsSafe();
            END_IF

            IF _pairs[1].SafeStateRequested THEN
                _funcTested[1] := TRUE;
            END_IF

            IF _pairs[2].SafeStateRequested THEN
                _funcTested[2] := TRUE;
            END_IF

            IF (NOT _pairs[1].IsActive OR _funcTested[1]) AND (NOT _pairs[2].IsActive OR _funcTested[2]) THEN
                _state := E_SafeMonState.Safe;
            END_IF

        E_SafeMonState.Safe:
            IF StateChanged() THEN
                SetOutputsSafe();
                _delayRunning := FALSE;
            END_IF

            IF _restartConnected THEN
                IF Restart THEN
                    IF NOT EdmInputsOk() THEN
                        _state := E_SafeMonState.Error;
                    ELSIF NOT safeRequested THEN
                        _state := E_SafeMonState.Start;
                    END_IF
                END_IF
            ELSIF NOT safeRequested AND EdmInputsTrue() THEN
                // automatic restart: an EDM fault keeps the FB in SAFE without an error
                _state := E_SafeMonState.Run;
            END_IF

        E_SafeMonState.Start:
            IF StateChanged() THEN
                SetOutputsSafe();
            END_IF

            IF safeRequested THEN
                _state := E_SafeMonState.Safe;
            ELSIF restartFalling THEN
                IF EdmInputsOk() THEN
                    _state := E_SafeMonState.Run;
                ELSE
                    _state := E_SafeMonState.Error;
                END_IF
            END_IF

        E_SafeMonState.Run:
            IF StateChanged() THEN
                MonOut    := TRUE;
                MonDelOut := TRUE;
                StartEdmResetMonitoring();
            END_IF

            IF NOT EdmResetOk() THEN
                _state := E_SafeMonState.Error;
            ELSIF safeRequested THEN
                IF Parameters.DelayTime > T#0S THEN
                    _state := E_SafeMonState.DelayOut;
                ELSE
                    _state := E_SafeMonState.Safe;
                END_IF
            END_IF

        E_SafeMonState.DelayOut:
            IF StateChanged() THEN
                MonOut    := FALSE;
                MonDelOut := TRUE;
                _delayTimer(IN := FALSE, PT := Parameters.DelayTime);
                _delayRunning := TRUE;
            END_IF

            _delayTimer(IN := TRUE, PT := Parameters.DelayTime);

            IF _delayTimer.Q THEN
                _state := E_SafeMonState.Safe;
            END_IF

        E_SafeMonState.ErrorDelay:
            IF StateChanged() THEN
                MonOut    := FALSE;
                MonDelOut := TRUE;

                IF NOT _delayRunning THEN
                    _delayTimer(IN := FALSE, PT := Parameters.DelayTime);
                    _delayRunning := TRUE;
                END_IF
            END_IF

            _delayTimer(IN := TRUE, PT := Parameters.DelayTime);

            IF _delayTimer.Q THEN
                _state := E_SafeMonState.Error;
            END_IF

        E_SafeMonState.Error:
            IF StateChanged() THEN
                SetOutputsSafe();
                Error         := TRUE;
                _delayRunning := FALSE;
            END_IF

            UpdateDiscrepancyDiag();

            IF _errAck AND NOT discError THEN
                _state := E_SafeMonState.Reset;
            END_IF

        E_SafeMonState.Reset:
            IF StateChanged() THEN
                SetOutputsSafe();
                Error := FALSE;
                Diag  := 0;
            END_IF

            IF _errAckFallingEdge THEN
                _state := SEL(_fbRun, E_SafeMonState.Stop, E_SafeMonState.Safe);
            END_IF
    END_CASE

    passes := passes + 1;
UNTIL (stateBefore = _state) OR (passes >= 3)
END_REPEAT

State := TO_BYTE(_state);
END_METHOD

METHOD PRIVATE SetOutputsSafe
MonOut    := FALSE;
MonDelOut := FALSE;
END_METHOD

METHOD PRIVATE StartEdmResetMonitoring
_edm1Dropped := FALSE;
_edm2Dropped := FALSE;
_edmResetTimer1(IN := FALSE, PT := Parameters.Edm1ResetTime);
_edmResetTimer2(IN := FALSE, PT := Parameters.Edm2ResetTime);
END_METHOD

METHOD PRIVATE StateChanged : BOOL
IF _prevState = _state THEN
    RETURN;
END_IF

_prevState   := _state;
StateChanged := TRUE;
END_METHOD

// Mirrors the discrepancy state of every pair into the diagnostic bits.
METHOD PRIVATE UpdateDiscrepancyDiag
VAR
    i : USINT;
END_VAR
FOR i := 1 TO 3 DO
    IF _pairs[i].DiscrepancyError THEN
        SetDiagBit(i - 1);

        IF _pairs[i].AwaitingSafeInputs THEN
            SetDiagBit(i + 7);
        ELSE
            ClearDiagBit(i + 7);
        END_IF
    END_IF
END_FOR
END_METHOD

END_FUNCTION_BLOCK

// ---- Tests/T_SafeTwoHand_Tests.TcPOU
FUNCTION_BLOCK T_SafeTwoHand_Tests EXTENDS TcUnit.FB_TestSuite
VAR
    // Test_BothHandsGiveOutputAndReleaseNeedsBothOff
    group_1 : T_SafeGroup;
    fb_1 : T_SafeTwoHand(group := group_1);
    // Test_SecondHandWithoutFirstGivesTwoHandError
    group_2 : T_SafeGroup;
    fb_2 : T_SafeTwoHand(group := group_2);
    // Test_HandDiscrepancyTimeout
    group_3 : T_SafeGroup;
    // SafeInputsAfterDiscError TRUE (not the default) so the error waits for both hands released (diag bit 10)
    fb_3 : T_SafeTwoHand(group := group_3) := (Parameters := (HandDiscrepancyTime := T#100MS, SafeInputsAfterDiscError := TRUE));
    state_3 : INT := 10;
    waitTimer_3 : TON;
END_VAR

Test_BothHandsGiveOutputAndReleaseNeedsBothOff();
Test_SecondHandWithoutFirstGivesTwoHandError();
Test_HandDiscrepancyTimeout();

METHOD PRIVATE Test_BothHandsGiveOutputAndReleaseNeedsBothOff
TcUnit.TEST(__POUNAME());
// arrange: single channel per hand
group_1(Run := TRUE);
fb_1(Twohand1 := FALSE, Twohand3 := FALSE);
// act
group_1(Run := TRUE);
fb_1(Twohand1 := TRUE, Twohand3 := FALSE);
AssertEquals_BYTE(Expected := TO_BYTE(E_SafeTwoHandState.OneButton), Actual := fb_1.State, Message := 'state 1BUTTON');
group_1(Run := TRUE);
fb_1(Twohand1 := TRUE, Twohand3 := TRUE);
// assert
AssertEquals_BOOL(Expected := TRUE, Actual := fb_1.TwoHandOut, Message := 'output on with both hands');
group_1(Run := TRUE);
fb_1(Twohand1 := FALSE, Twohand3 := TRUE);
AssertEquals_BOOL(Expected := FALSE, Actual := fb_1.TwoHandOut, Message := 'output off when one hand released');
AssertEquals_BYTE(Expected := TO_BYTE(E_SafeTwoHandState.Release), Actual := fb_1.State, Message := 'state RELEASE');
group_1(Run := TRUE);
fb_1(Twohand1 := TRUE, Twohand3 := TRUE);
AssertEquals_BOOL(Expected := FALSE, Actual := fb_1.TwoHandOut, Message := 'no re-trigger until both hands released');
TEST_FINISHED_NAMED(__POUNAME());
END_METHOD

METHOD PRIVATE Test_HandDiscrepancyTimeout
TcUnit.TEST(__POUNAME());
waitTimer_3();

CASE state_3 OF
    10:
        group_3(Run := TRUE);
        fb_3(Twohand1 := FALSE, Twohand3 := FALSE);
        state_3 := 20;
        waitTimer_3(IN := TRUE, PT := T#250MS);
    20:
        // act: only one hand for longer than the discrepancy time
        group_3(Run := TRUE);
        fb_3(Twohand1 := TRUE, Twohand3 := FALSE);

        IF NOT waitTimer_3.Q THEN
            RETURN;
        END_IF

        waitTimer_3(IN := FALSE);
        // assert
        AssertEquals_BOOL(Expected := TRUE, Actual := fb_3.Error, Message := 'discrepancy error between hands');
        AssertEquals_WORD(Expected := WORD#16#0404, Actual := fb_3.Diag, Message := 'diag bits 2 and 10');
        TEST_FINISHED_NAMED(__POUNAME());
        state_3 := 10;
END_CASE
END_METHOD

METHOD PRIVATE Test_SecondHandWithoutFirstGivesTwoHandError
TcUnit.TEST(__POUNAME());
// arrange
group_2(Run := TRUE);
fb_2(Twohand1 := FALSE, Twohand3 := FALSE);
group_2(Run := TRUE);
fb_2(Twohand1 := TRUE, Twohand3 := FALSE);
// act: first hand lost as the second is actuated
group_2(Run := TRUE);
fb_2(Twohand1 := FALSE, Twohand3 := TRUE);
// assert
AssertEquals_BOOL(Expected := TRUE, Actual := fb_2.Error, Message := 'two-hand error');
AssertEquals_WORD(Expected := WORD#64, Actual := fb_2.Diag, Message := 'diag bit 6');
TEST_FINISHED_NAMED(__POUNAME());
END_METHOD

END_FUNCTION_BLOCK

// ---- FunctionBlocks/T_SafeTwoHand.TcPOU
// Model of the TwinSAFE FB TWOHAND (two-hand control).
// Both hands (input pairs) must be actuated, optionally within HandDiscrepancyTime of each other.
// The output can only be set again after both hands were released together.
{attribute 'reflection'}
FUNCTION_BLOCK T_SafeTwoHand EXTENDS T_SafeFunctionBlockBase
VAR_INPUT
    Twohand1 : BOOL; // first hand, channel 1
    Twohand2 : BOOL; // first hand, channel 2
    Twohand3 : BOOL; // second hand, channel 1
    Twohand4 : BOOL; // second hand, channel 2
    Parameters : ST_SafeTwoHandParameters;
END_VAR
VAR_OUTPUT
    TwoHandOut : BOOL;
END_VAR
VAR
    {attribute 'is_connected' := 'Twohand1'}
    _twohand1Connected : BOOL;
    {attribute 'is_connected' := 'Twohand2'}
    _twohand2Connected : BOOL;
    {attribute 'is_connected' := 'Twohand3'}
    _twohand3Connected : BOOL;
    {attribute 'is_connected' := 'Twohand4'}
    _twohand4Connected : BOOL;
    _pairs : ARRAY[1..2] OF T_SafeInputPair;
    _state : E_SafeTwoHandState := E_SafeTwoHandState.Stop;
    _prevState : E_SafeTwoHandState;
    _handTimer : TON;
    _awaitingRelease : BOOL; // between-hands discrepancy error waits for both hands released
END_VAR

SUPER^();

METHOD PROTECTED Process
VAR
    acknowledge : BOOL;
    hand1 : BOOL; // first hand fully actuated
    hand2 : BOOL; // second hand fully actuated
    anyFalse : BOOL; // at least one active input released
    allFalse : BOOL; // every active input released
    discError : BOOL;
    operating : BOOL;
    stateBefore : E_SafeTwoHandState;
    passes : USINT;
END_VAR
acknowledge := (_state = E_SafeTwoHandState.Error) AND _errAck AND NOT _awaitingRelease;
_pairs[1](
    In1 := Twohand1,
    In2 := Twohand2,
    Active1 := _twohand1Connected,
    Active2 := _twohand2Connected,
    MakeContact1 := Parameters.Twohand1MakeContact,
    MakeContact2 := Parameters.Twohand2MakeContact,
    DiscrepancyTime := Parameters.DiscrepancyTime1,
    Monitor := _fbRun,
    SafeInputsAfterDiscError := Parameters.SafeInputsAfterDiscError,
    Acknowledge := acknowledge
);

_pairs[2](
    In1 := Twohand3,
    In2 := Twohand4,
    Active1 := _twohand3Connected,
    Active2 := _twohand4Connected,
    MakeContact1 := Parameters.Twohand3MakeContact,
    MakeContact2 := Parameters.Twohand4MakeContact,
    DiscrepancyTime := Parameters.DiscrepancyTime2,
    Monitor := _fbRun,
    SafeInputsAfterDiscError := Parameters.SafeInputsAfterDiscError,
    Acknowledge := acknowledge
);

hand1     := _pairs[1].IsActive AND _pairs[1].AllTrue;
hand2     := _pairs[2].IsActive AND _pairs[2].AllTrue;
anyFalse  := NOT (_pairs[1].AllTrue AND _pairs[2].AllTrue);
allFalse  := (NOT _pairs[1].IsActive OR _pairs[1].AllFalse) AND (NOT _pairs[2].IsActive OR _pairs[2].AllFalse);
discError := _pairs[1].DiscrepancyError OR _pairs[2].DiscrepancyError;

IF NOT _fbRun AND _state <> E_SafeTwoHandState.Error AND _state <> E_SafeTwoHandState.Reset THEN
    _state := E_SafeTwoHandState.Stop;
END_IF

operating := (_state = E_SafeTwoHandState.Safe)
                 OR (_state = E_SafeTwoHandState.OneButton)
                 OR (_state = E_SafeTwoHandState.TwoButton)
                 OR (_state = E_SafeTwoHandState.Run)
                 OR (_state = E_SafeTwoHandState.Release);

IF discError AND operating THEN
    UpdateDiscrepancyDiag();
    _state := E_SafeTwoHandState.Error;
END_IF

IF _awaitingRelease AND allFalse THEN
    _awaitingRelease := FALSE;
END_IF

passes := 0;

REPEAT
    stateBefore := _state;

    CASE _state OF
        E_SafeTwoHandState.Stop:
            IF StateChanged() THEN
                TwoHandOut := FALSE;
                Error      := FALSE;
                Diag       := 0;
            END_IF

            IF _fbRun THEN
                _state := E_SafeTwoHandState.Safe;
            END_IF

        E_SafeTwoHandState.Safe:
            IF StateChanged() THEN
                TwoHandOut := FALSE;
            END_IF

            IF hand1 THEN
                _state := E_SafeTwoHandState.OneButton;
            ELSIF hand2 THEN
                _state := E_SafeTwoHandState.TwoButton;
            END_IF

        E_SafeTwoHandState.OneButton:
            IF StateChanged() THEN
                _handTimer(IN := FALSE, PT := Parameters.HandDiscrepancyTime);
            END_IF

            _handTimer(IN := (Parameters.HandDiscrepancyTime > T#0S), PT := Parameters.HandDiscrepancyTime);

            IF _handTimer.Q THEN
                SetHandDiscrepancyError();
            ELSIF hand1 AND hand2 THEN
                _state := E_SafeTwoHandState.Run;
            ELSIF hand2 THEN
                // second hand actuated while the first is no longer detected
                SetDiagBit(6);
                _state := E_SafeTwoHandState.Error;
            ELSIF NOT hand1 THEN
                _state := SEL(allFalse, E_SafeTwoHandState.Release, E_SafeTwoHandState.Safe);
            END_IF

        E_SafeTwoHandState.TwoButton:
            IF StateChanged() THEN
                _handTimer(IN := FALSE, PT := Parameters.HandDiscrepancyTime);
            END_IF

            _handTimer(IN := (Parameters.HandDiscrepancyTime > T#0S), PT := Parameters.HandDiscrepancyTime);

            IF _handTimer.Q THEN
                SetHandDiscrepancyError();
            ELSIF hand1 AND hand2 THEN
                _state := E_SafeTwoHandState.Run;
            ELSIF hand1 THEN
                SetDiagBit(6);
                _state := E_SafeTwoHandState.Error;
            ELSIF NOT hand2 THEN
                _state := SEL(allFalse, E_SafeTwoHandState.Release, E_SafeTwoHandState.Safe);
            END_IF

        E_SafeTwoHandState.Run:
            IF StateChanged() THEN
                TwoHandOut := TRUE;
            END_IF

            IF anyFalse THEN
                _state := E_SafeTwoHandState.Release;
            END_IF

        E_SafeTwoHandState.Release:
            IF StateChanged() THEN
                TwoHandOut := FALSE;
            END_IF

            IF allFalse THEN
                _state := E_SafeTwoHandState.Safe;
            END_IF

        E_SafeTwoHandState.Error:
            IF StateChanged() THEN
                TwoHandOut := FALSE;
                Error      := TRUE;
            END_IF

            UpdateDiscrepancyDiag();

            IF _awaitingRelease THEN
                SetDiagBit(10);
            ELSE
                ClearDiagBit(10);
            END_IF

            IF _errAck AND NOT _awaitingRelease AND NOT discError THEN
                _state := E_SafeTwoHandState.Reset;
            END_IF

        E_SafeTwoHandState.Reset:
            IF StateChanged() THEN
                TwoHandOut := FALSE;
                Error      := FALSE;
                Diag       := 0;
            END_IF

            IF _errAckFallingEdge THEN
                _state := SEL(_fbRun, E_SafeTwoHandState.Stop, E_SafeTwoHandState.Safe);
            END_IF
    END_CASE

    passes := passes + 1;
UNTIL (stateBefore = _state) OR (passes >= 3)
END_REPEAT

State := TO_BYTE(_state);
END_METHOD

METHOD PRIVATE SetHandDiscrepancyError
SetDiagBit(2);
_awaitingRelease := Parameters.SafeInputsAfterDiscError;
_state           := E_SafeTwoHandState.Error;
END_METHOD

METHOD PRIVATE StateChanged : BOOL
IF _prevState = _state THEN
    RETURN;
END_IF

_prevState   := _state;
StateChanged := TRUE;
END_METHOD

PROPERTY TwoHandState : E_SafeTwoHandState
GET
TwoHandState := _state;
END_GET
END_PROPERTY

// Mirrors the discrepancy state of every pair into the diagnostic bits.
METHOD PRIVATE UpdateDiscrepancyDiag
VAR
    i : USINT;
END_VAR
FOR i := 1 TO 2 DO
    IF _pairs[i].DiscrepancyError THEN
        SetDiagBit(i - 1);

        IF _pairs[i].AwaitingSafeInputs THEN
            SetDiagBit(i + 7);
        ELSE
            ClearDiagBit(i + 7);
        END_IF
    END_IF
END_FOR
END_METHOD

END_FUNCTION_BLOCK

// ---- Tests/T_SafeMuting_Tests.TcPOU
FUNCTION_BLOCK T_SafeMuting_Tests EXTENDS TcUnit.FB_TestSuite
VAR
    // Test_OssdBlockedWithoutMutingGivesSafe
    group_1 : T_SafeGroup;
    fb_1 : T_SafeMuting(group := group_1);
    // Test_SequentialMutingKeepsOutputOn
    group_2 : T_SafeGroup;
    fb_2 : T_SafeMuting(group := group_2) := (Parameters := (SequentialInputs := TRUE));
    // Test_SequenceViolationGivesError
    group_3 : T_SafeGroup;
    fb_3 : T_SafeMuting(group := group_3) := (Parameters := (SequentialInputs := TRUE));
    // Test_TwoSensorParallelSequence
    group_4 : T_SafeGroup;
    fb_4 : T_SafeMuting(group := group_4);
    // Test_ResetTimeNotMultipleOfTenIsRefused
    group_5 : T_SafeGroup;
    fb_5 : T_SafeMuting(group := group_5) := (Parameters := (Edm1ResetTime := T#25MS));
END_VAR

Test_OssdBlockedWithoutMutingGivesSafe();
Test_SequentialMutingKeepsOutputOn();
Test_SequenceViolationGivesError();
Test_TwoSensorParallelSequence();
Test_ResetTimeNotMultipleOfTenIsRefused();

METHOD PRIVATE Test_OssdBlockedWithoutMutingGivesSafe
TcUnit.TEST(__POUNAME());
// arrange: only the protective device connected
group_1(Run := TRUE);
fb_1(OSSDIn1 := TRUE);
group_1(Run := TRUE);
fb_1(OSSDIn1 := TRUE);
AssertEquals_BOOL(Expected := TRUE, Actual := fb_1.MuteOut, Message := 'output on with clear protective device');
// act
group_1(Run := TRUE);
fb_1(OSSDIn1 := FALSE);
// assert
AssertEquals_BOOL(Expected := FALSE, Actual := fb_1.MuteOut, Message := 'output off when interrupted');
AssertEquals_BYTE(Expected := TO_BYTE(E_SafeMutingState.Safe), Actual := fb_1.State, Message := 'state SAFE');
group_1(Run := TRUE);
fb_1(OSSDIn1 := TRUE);
AssertEquals_BOOL(Expected := TRUE, Actual := fb_1.MuteOut, Message := 'automatic restart when clear again');
TEST_FINISHED_NAMED(__POUNAME());
END_METHOD

METHOD PRIVATE Test_SequenceViolationGivesError
TcUnit.TEST(__POUNAME());
// arrange
group_3(Run := TRUE);
fb_3(
    MutingEnable := TRUE,
    MutingIn1 := FALSE,
    MutingIn2 := FALSE,
    MutingIn3 := FALSE,
    MutingIn4 := FALSE,
    OSSDIn1 := TRUE
);

group_3(Run := TRUE);
fb_3(
    MutingEnable := TRUE,
    MutingIn1 := FALSE,
    MutingIn2 := FALSE,
    MutingIn3 := FALSE,
    MutingIn4 := FALSE,
    OSSDIn1 := TRUE
);

group_3(Run := TRUE);
fb_3(
    MutingEnable := TRUE,
    MutingIn1 := TRUE,
    MutingIn2 := FALSE,
    MutingIn3 := FALSE,
    MutingIn4 := FALSE,
    OSSDIn1 := TRUE
);

// act: OSSD blocked before the second sensor
group_3(Run := TRUE);
fb_3(
    MutingEnable := TRUE,
    MutingIn1 := TRUE,
    MutingIn2 := FALSE,
    MutingIn3 := FALSE,
    MutingIn4 := FALSE,
    OSSDIn1 := FALSE
);

// assert
AssertEquals_BOOL(Expected := TRUE, Actual := fb_3.Error, Message := 'sequence violation');
AssertEquals_WORD(Expected := WORD#64, Actual := fb_3.Diag, Message := 'diag bit 6');
AssertEquals_BOOL(Expected := FALSE, Actual := fb_3.MuteOut, Message := 'output off');
TEST_FINISHED_NAMED(__POUNAME());
END_METHOD

METHOD PRIVATE Test_SequentialMutingKeepsOutputOn
TcUnit.TEST(__POUNAME());
// arrange: four single-channel sensors, running
group_2(Run := TRUE);
fb_2(
    MutingEnable := TRUE,
    MutingIn1 := FALSE,
    MutingIn2 := FALSE,
    MutingIn3 := FALSE,
    MutingIn4 := FALSE,
    OSSDIn1 := TRUE
);

group_2(Run := TRUE);
fb_2(
    MutingEnable := TRUE,
    MutingIn1 := FALSE,
    MutingIn2 := FALSE,
    MutingIn3 := FALSE,
    MutingIn4 := FALSE,
    OSSDIn1 := TRUE
);

// act: M1, M2, OSSD blocked, M3, M1 off, M4, M2 off, OSSD clear, M3 off, M4 off
group_2(Run := TRUE);
fb_2(
    MutingEnable := TRUE,
    MutingIn1 := TRUE,
    MutingIn2 := FALSE,
    MutingIn3 := FALSE,
    MutingIn4 := FALSE,
    OSSDIn1 := TRUE
);

AssertEquals_BYTE(Expected := TO_BYTE(E_SafeMutingState.Muting1), Actual := fb_2.State, Message := 'MUTING1');
AssertEquals_BOOL(Expected := TRUE, Actual := fb_2.MutingActive, Message := 'muting active');
group_2(Run := TRUE);
fb_2(
    MutingEnable := TRUE,
    MutingIn1 := TRUE,
    MutingIn2 := TRUE,
    MutingIn3 := FALSE,
    MutingIn4 := FALSE,
    OSSDIn1 := TRUE
);

group_2(Run := TRUE);
fb_2(
    MutingEnable := TRUE,
    MutingIn1 := TRUE,
    MutingIn2 := TRUE,
    MutingIn3 := FALSE,
    MutingIn4 := FALSE,
    OSSDIn1 := FALSE
);

AssertEquals_BYTE(Expected := TO_BYTE(E_SafeMutingState.Muting3), Actual := fb_2.State, Message := 'MUTING3');
AssertEquals_BOOL(Expected := TRUE, Actual := fb_2.MuteOut, Message := 'output stays on while muted');
group_2(Run := TRUE);
fb_2(
    MutingEnable := TRUE,
    MutingIn1 := TRUE,
    MutingIn2 := TRUE,
    MutingIn3 := TRUE,
    MutingIn4 := FALSE,
    OSSDIn1 := FALSE
);

group_2(Run := TRUE);
fb_2(
    MutingEnable := TRUE,
    MutingIn1 := FALSE,
    MutingIn2 := TRUE,
    MutingIn3 := TRUE,
    MutingIn4 := FALSE,
    OSSDIn1 := FALSE
);

group_2(Run := TRUE);
fb_2(
    MutingEnable := TRUE,
    MutingIn1 := FALSE,
    MutingIn2 := TRUE,
    MutingIn3 := TRUE,
    MutingIn4 := TRUE,
    OSSDIn1 := FALSE
);

group_2(Run := TRUE);
fb_2(
    MutingEnable := TRUE,
    MutingIn1 := FALSE,
    MutingIn2 := FALSE,
    MutingIn3 := TRUE,
    MutingIn4 := TRUE,
    OSSDIn1 := FALSE
);

group_2(Run := TRUE);
fb_2(
    MutingEnable := TRUE,
    MutingIn1 := FALSE,
    MutingIn2 := FALSE,
    MutingIn3 := TRUE,
    MutingIn4 := TRUE,
    OSSDIn1 := TRUE
);

AssertEquals_BYTE(Expected := TO_BYTE(E_SafeMutingState.Muting8), Actual := fb_2.State, Message := 'MUTING8');
group_2(Run := TRUE);
fb_2(
    MutingEnable := TRUE,
    MutingIn1 := FALSE,
    MutingIn2 := FALSE,
    MutingIn3 := FALSE,
    MutingIn4 := TRUE,
    OSSDIn1 := TRUE
);

group_2(Run := TRUE);
fb_2(
    MutingEnable := TRUE,
    MutingIn1 := FALSE,
    MutingIn2 := FALSE,
    MutingIn3 := FALSE,
    MutingIn4 := FALSE,
    OSSDIn1 := TRUE
);

// assert
AssertEquals_BYTE(Expected := TO_BYTE(E_SafeMutingState.Run), Actual := fb_2.State, Message := 'RUN after the sequence');
AssertEquals_BOOL(Expected := FALSE, Actual := fb_2.MutingActive, Message := 'muting no longer active');
AssertEquals_BOOL(Expected := FALSE, Actual := fb_2.Error, Message := 'no error');
TEST_FINISHED_NAMED(__POUNAME());
END_METHOD

METHOD PRIVATE Test_TwoSensorParallelSequence
TcUnit.TEST(__POUNAME());
// arrange: two two-channel sensors (parallel inputs), running
group_4(Run := TRUE);
fb_4(
    MutingEnable := TRUE,
    MutingIn1 := FALSE,
    MutingIn2 := FALSE,
    MutingIn3 := FALSE,
    MutingIn4 := FALSE,
    OSSDIn1 := TRUE
);

group_4(Run := TRUE);
fb_4(
    MutingEnable := TRUE,
    MutingIn1 := FALSE,
    MutingIn2 := FALSE,
    MutingIn3 := FALSE,
    MutingIn4 := FALSE,
    OSSDIn1 := TRUE
);

// act: S1, S2, OSSD blocked, S1 off, OSSD clear, S2 off
group_4(Run := TRUE);
fb_4(
    MutingEnable := TRUE,
    MutingIn1 := TRUE,
    MutingIn2 := TRUE,
    MutingIn3 := FALSE,
    MutingIn4 := FALSE,
    OSSDIn1 := TRUE
);

group_4(Run := TRUE);
fb_4(
    MutingEnable := TRUE,
    MutingIn1 := TRUE,
    MutingIn2 := TRUE,
    MutingIn3 := TRUE,
    MutingIn4 := TRUE,
    OSSDIn1 := TRUE
);

group_4(Run := TRUE);
fb_4(
    MutingEnable := TRUE,
    MutingIn1 := TRUE,
    MutingIn2 := TRUE,
    MutingIn3 := TRUE,
    MutingIn4 := TRUE,
    OSSDIn1 := FALSE
);

AssertEquals_BOOL(Expected := TRUE, Actual := fb_4.MuteOut, Message := 'output stays on while muted');
group_4(Run := TRUE);
fb_4(
    MutingEnable := TRUE,
    MutingIn1 := FALSE,
    MutingIn2 := FALSE,
    MutingIn3 := TRUE,
    MutingIn4 := TRUE,
    OSSDIn1 := FALSE
);

group_4(Run := TRUE);
fb_4(
    MutingEnable := TRUE,
    MutingIn1 := FALSE,
    MutingIn2 := FALSE,
    MutingIn3 := TRUE,
    MutingIn4 := TRUE,
    OSSDIn1 := TRUE
);

group_4(Run := TRUE);
fb_4(
    MutingEnable := TRUE,
    MutingIn1 := FALSE,
    MutingIn2 := FALSE,
    MutingIn3 := FALSE,
    MutingIn4 := FALSE,
    OSSDIn1 := TRUE
);

// assert
AssertEquals_BYTE(Expected := TO_BYTE(E_SafeMutingState.Run), Actual := fb_4.State, Message := 'RUN after the sequence');
AssertEquals_BOOL(Expected := FALSE, Actual := fb_4.Error, Message := 'no error');
TEST_FINISHED_NAMED(__POUNAME());
END_METHOD

METHOD PRIVATE Test_ResetTimeNotMultipleOfTenIsRefused
TcUnit.TEST(__POUNAME());
// arrange / act: Edm1ResetTime is 25 ms, which the Safety Editor refuses
group_5(Run := TRUE);
fb_5(EDM1 := TRUE, OSSDIn1 := TRUE);
group_5(Run := TRUE);
fb_5(EDM1 := TRUE, OSSDIn1 := TRUE);
// assert
AssertEquals_BOOL(Expected := TRUE, Actual := fb_5.Error, Message := 'configuration error reported');
AssertEquals_BYTE(Expected := TO_BYTE(E_SafeFbState.Error), Actual := fb_5.State, Message := 'state ERROR');
AssertEquals_WORD(Expected := WORD#16#8000, Actual := fb_5.Diag, Message := 'diag bit 15 configuration refused');
AssertEquals_BOOL(Expected := FALSE, Actual := fb_5.MuteOut, Message := 'MuteOut stays at its safe value');
AssertEquals_BOOL(Expected := TRUE, Actual := group_5.FbErr, Message := 'the group sees an FB error');
// act: ErrAck 0 -> 1 -> 0 does not clear a configuration error
group_5(Run := TRUE, ErrAck := TRUE);
fb_5(EDM1 := TRUE, OSSDIn1 := TRUE);
group_5(Run := TRUE, ErrAck := TRUE);
fb_5(EDM1 := TRUE, OSSDIn1 := TRUE);
group_5(Run := TRUE, ErrAck := FALSE);
fb_5(EDM1 := TRUE, OSSDIn1 := TRUE);
AssertEquals_BOOL(Expected := TRUE, Actual := fb_5.Error, Message := 'error not acknowledged');
AssertEquals_WORD(Expected := WORD#16#8000, Actual := fb_5.Diag, Message := 'diag bit 15 kept');
TEST_FINISHED_NAMED(__POUNAME());
END_METHOD

END_FUNCTION_BLOCK

// ---- FunctionBlocks/T_SafeMuting.TcPOU
// Model of the TwinSAFE FB MUTING.
// Suppresses the protective device (OSSDIn) while the muting sensors are actuated in the expected order.
// Sequence (sequential inputs, four sensors, forward):
//   M1 on, M2 on, OSSD blocked, M3 on, M1 off, M4 on, M2 off, OSSD clear, M3 off, M4 off
// Sequence (two sensors: parallel inputs, or sequential with MutingIn3/4 unconnected):
//   S1 on, S2 on, OSSD blocked, S1 off, OSSD clear, S2 off
// Any other change of a sensor or the OSSD during a sequence violates it (diagnostic bit 6).
// The Safety Editor refuses an EDM reset time that is not 0 ms, a multiple of 10 ms and at most 60000 ms:
// the model then reports Error with diagnostic bit 15 instead of running (see T_SafeFunctionBlockBase).
{attribute 'reflection'}
FUNCTION_BLOCK T_SafeMuting EXTENDS T_SafeFunctionBlockBase
VAR_INPUT
    MutingEnable : BOOL; // may be a standard PLC signal
    EDM1 : BOOL; // feedback loop of MuteOut
    EDM2 : BOOL; // feedback loop of MuteDelOut
    MutingIn1 : BOOL;
    MutingIn2 : BOOL;
    OSSDIn1 : BOOL; // protective device channel 1 (TRUE = clear)
    OSSDIn2 : BOOL; // protective device channel 2
    MutingIn3 : BOOL;
    MutingIn4 : BOOL;
    Parameters : ST_SafeMutingParameters;
END_VAR
VAR_OUTPUT
    MutingActive : BOOL; // muting lamp
    MuteOut : BOOL;
    MuteDelOut : BOOL;
END_VAR
VAR
    {attribute 'is_connected' := 'MutingEnable'}
    _mutingEnableConnected : BOOL;
    {attribute 'is_connected' := 'EDM1'}
    _eDM1Connected : BOOL;
    {attribute 'is_connected' := 'EDM2'}
    _eDM2Connected : BOOL;
    {attribute 'is_connected' := 'MutingIn1'}
    _mutingIn1Connected : BOOL;
    {attribute 'is_connected' := 'MutingIn2'}
    _mutingIn2Connected : BOOL;
    {attribute 'is_connected' := 'OSSDIn1'}
    _oSSDIn1Connected : BOOL;
    {attribute 'is_connected' := 'OSSDIn2'}
    _oSSDIn2Connected : BOOL;
    {attribute 'is_connected' := 'MutingIn3'}
    _mutingIn3Connected : BOOL;
    {attribute 'is_connected' := 'MutingIn4'}
    _mutingIn4Connected : BOOL;
    _pairs : ARRAY[1..3] OF T_SafeInputPair; // 1: MutingIn1/2, 2: MutingIn3/4, 3: OSSDIn1/2
    _state : E_SafeMutingState := E_SafeMutingState.Stop;
    _prevState : E_SafeMutingState;
    _filterTimers : ARRAY[1..4] OF TON;
    _filtered : ARRAY[1..4] OF BOOL;
    _sensor : ARRAY[1..4] OF BOOL; // actuated sensors after configuration
    _ossdBlocked : BOOL;
    _sensorCount : USINT;
    _seqSensor : ARRAY[1..10] OF USINT; // 0 = OSSD
    _seqLevel : ARRAY[1..10] OF BOOL;
    _seqLength : USINT;
    _seqIndex : USINT; // consumed events
    _expected : ARRAY[0..4] OF BOOL; // expected level of each signal (0 = OSSD blocked)
    _maxTimer : TON;
    _delayTimer : TON;
    _pendingError : BOOL;
    _edmResetTimer1 : TON;
    _edmResetTimer2 : TON;
    _edm1Dropped : BOOL;
    _edm2Dropped : BOOL;
END_VAR

SUPER^();

// The EDM reset times must be 0 ms or a multiple of 10 ms up to 60000 ms (Safety Editor: "'Reset Time' parameter ... has to be 0 ms or a multiple of 10 ms and maximal 60000 ms").
METHOD PROTECTED ConfigurationOk : BOOL
IF NOT F_SafeResetTimeOk(Parameters.Edm1ResetTime) THEN
    _configurationFault := 'T_SafeMuting: $'Reset Time$' parameter of EDM1 of MUTING has to be 0 ms or a multiple of 10 ms and maximal 60000 ms';
    RETURN;
ELSIF NOT F_SafeResetTimeOk(Parameters.Edm2ResetTime) THEN
    _configurationFault := 'T_SafeMuting: $'Reset Time$' parameter of EDM2 of MUTING has to be 0 ms or a multiple of 10 ms and maximal 60000 ms';
    RETURN;
END_IF

ConfigurationOk := TRUE;
END_METHOD

METHOD PRIVATE Actual : BOOL
VAR_INPUT
    signal : USINT; // 0 = OSSD blocked, 1..4 = sensor actuated
END_VAR
IF signal = 0 THEN
    Actual := _ossdBlocked;
ELSE
    Actual := _sensor[signal];
END_IF
END_METHOD

METHOD PRIVATE AddEvent
VAR_INPUT
    sensor : USINT; // 0 = OSSD
    level : BOOL; // sensor actuated / OSSD blocked
    backwards : BOOL;
END_VAR
IF sensor = 0 AND Parameters.OssdCheckOptional THEN
    RETURN;
END_IF

IF _seqLength >= 10 THEN
    RETURN;
END_IF

_seqLength := _seqLength + 1;

IF sensor > 0 AND backwards THEN
    _seqSensor[_seqLength] := _sensorCount + 1 - sensor;
ELSE
    _seqSensor[_seqLength] := sensor;
END_IF

_seqLevel[_seqLength] := level;
END_METHOD

// Consumes every expected event that has occurred, then checks that no signal deviates
// from the expected pattern. Returns TRUE when the sequence has been violated.
METHOD PRIVATE Advance : BOOL
VAR
    progressed : BOOL;
    next : USINT;
    k : USINT;
END_VAR
REPEAT
    progressed := FALSE;

    IF _seqIndex < _seqLength THEN
        next := _seqIndex + 1;

        IF Actual(_seqSensor[next]) = _seqLevel[next] THEN
            _expected[_seqSensor[next]] := _seqLevel[next];
            _seqIndex                   := next;
            progressed                  := TRUE;
        END_IF
    END_IF
UNTIL NOT progressed
END_REPEAT

FOR k := 0 TO _sensorCount DO
    IF k = 0 AND Parameters.OssdCheckOptional THEN
        CONTINUE;
    END_IF

    IF Actual(k) <> _expected[k] THEN
        Advance := TRUE;
    END_IF
END_FOR
END_METHOD

METHOD PRIVATE AnySensor : BOOL
VAR
    k : USINT;
END_VAR
FOR k := 1 TO _sensorCount DO
    AnySensor := AnySensor OR _sensor[k];
END_FOR
END_METHOD

// Builds the expected event list for the configured sensor arrangement.
METHOD PRIVATE BuildSequence
VAR_INPUT
    backwards : BOOL;
END_VAR
_seqLength := 0;

IF _sensorCount = 4 THEN
    AddEvent(1, TRUE, backwards);
    AddEvent(2, TRUE, backwards);
    AddEvent(0, TRUE, backwards);
    AddEvent(3, TRUE, backwards);
    AddEvent(1, FALSE, backwards);
    AddEvent(4, TRUE, backwards);
    AddEvent(2, FALSE, backwards);
    AddEvent(0, FALSE, backwards);
    AddEvent(3, FALSE, backwards);
    AddEvent(4, FALSE, backwards);
ELSE
    AddEvent(1, TRUE, backwards);
    AddEvent(2, TRUE, backwards);
    AddEvent(0, TRUE, backwards);
    AddEvent(1, FALSE, backwards);
    AddEvent(0, FALSE, backwards);
    AddEvent(2, FALSE, backwards);
END_IF
END_METHOD

// Checks the EDM inputs at restart and records diagnostic bits 4/5 on failure.
METHOD PRIVATE EdmInputsOk : BOOL
EdmInputsOk := TRUE;

IF _eDM1Connected AND NOT EDM1 THEN
    SetDiagBit(4);
    EdmInputsOk := FALSE;
END_IF

IF _eDM2Connected AND NOT EDM2 THEN
    SetDiagBit(5);
    EdmInputsOk := FALSE;
END_IF
END_METHOD

// TRUE when every connected EDM input reads 1 (contactors released).
METHOD PRIVATE EdmInputsTrue : BOOL
EdmInputsTrue := (NOT _eDM1Connected OR EDM1) AND (NOT _eDM2Connected OR EDM2);
END_METHOD

// EL6910 extension: after the outputs switch on, each connected EDM input must drop to FALSE
// within its Reset Time. Returns FALSE (and sets diagnostic bits 4/5) on timeout.
METHOD PRIVATE EdmResetOk : BOOL
EdmResetOk := TRUE;

IF _eDM1Connected AND Parameters.Edm1ResetTime > T#0S THEN
    IF NOT EDM1 THEN
        _edm1Dropped := TRUE;
    END_IF

    _edmResetTimer1(IN := NOT _edm1Dropped, PT := Parameters.Edm1ResetTime);

    IF _edmResetTimer1.Q THEN
        SetDiagBit(4);
        EdmResetOk := FALSE;
    END_IF
END_IF

IF _eDM2Connected AND Parameters.Edm2ResetTime > T#0S THEN
    IF NOT EDM2 THEN
        _edm2Dropped := TRUE;
    END_IF

    _edmResetTimer2(IN := NOT _edm2Dropped, PT := Parameters.Edm2ResetTime);

    IF _edmResetTimer2.Q THEN
        SetDiagBit(5);
        EdmResetOk := FALSE;
    END_IF
END_IF
END_METHOD

METHOD PRIVATE IsMuting : BOOL
IsMuting := (TO_BYTE(_state) >= TO_BYTE(E_SafeMutingState.Muting1)) AND (TO_BYTE(_state) <= TO_BYTE(E_SafeMutingState.Muting9));
END_METHOD

PROPERTY MutingState : E_SafeMutingState
GET
MutingState := _state;
END_GET
END_PROPERTY

// State code for the given number of consumed sequence events.
METHOD PRIVATE MutingStateFor : E_SafeMutingState
VAR_INPUT
    consumed : USINT;
END_VAR
CASE consumed OF
    1:
        MutingStateFor := E_SafeMutingState.Muting1;
    2:
        MutingStateFor := E_SafeMutingState.Muting2;
    3:
        MutingStateFor := E_SafeMutingState.Muting3;
    4:
        MutingStateFor := E_SafeMutingState.Muting4;
    5:
        MutingStateFor := E_SafeMutingState.Muting5;
    6:
        MutingStateFor := E_SafeMutingState.Muting6;
    7:
        MutingStateFor := E_SafeMutingState.Muting7;
    8:
        MutingStateFor := E_SafeMutingState.Muting8;
    9:
        MutingStateFor := E_SafeMutingState.Muting9;
ELSE
    MutingStateFor := E_SafeMutingState.Run;
END_CASE
END_METHOD

METHOD PROTECTED Process
VAR
    raw : ARRAY[1..4] OF BOOL;
    i : USINT;
    acknowledge : BOOL;
    discError : BOOL;
    operating : BOOL;
    startFwd : BOOL;
    startBwd : BOOL;
    k : USINT;
    stateBefore : E_SafeMutingState;
    passes : USINT;
END_VAR
// Debounce of the muting inputs
raw[1] := MutingIn1;
raw[2] := MutingIn2;
raw[3] := MutingIn3;
raw[4] := MutingIn4;

FOR i := 1 TO 4 DO
    _filterTimers[i](IN := (raw[i] <> _filtered[i]), PT := Parameters.FilterTime);

    IF _filterTimers[i].Q OR Parameters.FilterTime = T#0S THEN
        _filtered[i] := raw[i];
    END_IF
END_FOR

acknowledge := (_state = E_SafeMutingState.Error) AND _errAck;
_pairs[1](
    In1 := _filtered[1],
    In2 := _filtered[2],
    Active1 := _mutingIn1Connected,
    Active2 := _mutingIn2Connected,
    MakeContact1 := Parameters.MutingIn1MakeContact,
    MakeContact2 := Parameters.MutingIn2MakeContact,
    DiscrepancyTime := Parameters.MutingDiscrepancyTime1,
    Monitor := _fbRun AND NOT Parameters.SequentialInputs,
    SafeInputsAfterDiscError := Parameters.SafeInputsAfterDiscError,
    Acknowledge := acknowledge
);

_pairs[2](
    In1 := _filtered[3],
    In2 := _filtered[4],
    Active1 := _mutingIn3Connected,
    Active2 := _mutingIn4Connected,
    MakeContact1 := Parameters.MutingIn3MakeContact,
    MakeContact2 := Parameters.MutingIn4MakeContact,
    DiscrepancyTime := Parameters.MutingDiscrepancyTime2,
    Monitor := _fbRun AND NOT Parameters.SequentialInputs,
    SafeInputsAfterDiscError := Parameters.SafeInputsAfterDiscError,
    Acknowledge := acknowledge
);

_pairs[3](
    In1 := OSSDIn1,
    In2 := OSSDIn2,
    Active1 := _oSSDIn1Connected,
    Active2 := _oSSDIn2Connected,
    MakeContact1 := Parameters.OSSDIn1MakeContact,
    MakeContact2 := Parameters.OSSDIn2MakeContact,
    DiscrepancyTime := Parameters.OssdDiscrepancyTime,
    Monitor := _fbRun,
    SafeInputsAfterDiscError := Parameters.SafeInputsAfterDiscError,
    Acknowledge := acknowledge
);

IF Parameters.SequentialInputs THEN
    _sensorCount := SEL(_mutingIn3Connected OR _mutingIn4Connected, 2, 4);
    _sensor[1]   := F_SafeInputValue(_mutingIn1Connected, Parameters.MutingIn1MakeContact, _filtered[1]);
    _sensor[2]   := F_SafeInputValue(_mutingIn2Connected, Parameters.MutingIn2MakeContact, _filtered[2]);
    _sensor[3]   := F_SafeInputValue(_mutingIn3Connected, Parameters.MutingIn3MakeContact, _filtered[3]);
    _sensor[4]   := F_SafeInputValue(_mutingIn4Connected, Parameters.MutingIn4MakeContact, _filtered[4]);
ELSE
    _sensorCount := 2;
    _sensor[1]   := _pairs[1].IsActive AND _pairs[1].AllTrue;
    _sensor[2]   := _pairs[2].IsActive AND _pairs[2].AllTrue;
    _sensor[3]   := FALSE;
    _sensor[4]   := FALSE;
END_IF

_ossdBlocked := NOT _pairs[3].AllTrue;

FOR i := 1 TO 3 DO
    discError := discError OR _pairs[i].DiscrepancyError;
END_FOR

IF NOT _fbRun AND _state <> E_SafeMutingState.Error AND _state <> E_SafeMutingState.Reset THEN
    _state := E_SafeMutingState.Stop;
END_IF

operating := (_state = E_SafeMutingState.Safe) OR (_state = E_SafeMutingState.Run) OR IsMuting();

IF discError THEN
    IF operating THEN
        UpdateDiscrepancyDiag();
        _state := E_SafeMutingState.Error;
    ELSIF _state = E_SafeMutingState.DelayOut THEN
        UpdateDiscrepancyDiag();
        _pendingError := TRUE;
    END_IF
END_IF

passes := 0;

REPEAT
    stateBefore := _state;

    CASE _state OF
        E_SafeMutingState.Stop:
            IF StateChanged() THEN
                SetOutputsSafe();
                MutingActive  := FALSE;
                Error         := FALSE;
                Diag          := 0;
                _pendingError := FALSE;
            END_IF

            IF _fbRun THEN
                _state := E_SafeMutingState.Safe;
            END_IF

        E_SafeMutingState.Safe:
            IF StateChanged() THEN
                SetOutputsSafe();
                MutingActive := FALSE;
            END_IF

            IF NOT _ossdBlocked AND EdmInputsTrue() THEN
                _state := E_SafeMutingState.Run;
            END_IF

        E_SafeMutingState.Run:
            IF StateChanged() THEN
                MuteOut      := TRUE;
                MuteDelOut   := TRUE;
                MutingActive := FALSE;
                StartEdmResetMonitoring();
                _seqIndex := 0;
                _maxTimer(IN := FALSE, PT := Parameters.MaxMutingTime);
            END_IF

            startFwd := _sensor[1];
            startBwd := Parameters.BackwardsMode AND _sensor[_sensorCount];

            IF NOT EdmResetOk() THEN
                _state := E_SafeMutingState.Error;
            ELSIF MutingEnable AND (startFwd OR startBwd) THEN
                BuildSequence(startBwd AND NOT startFwd);

                FOR k := 0 TO 4 DO
                    _expected[k] := FALSE;
                END_FOR

                _seqIndex := 0;

                IF Advance() THEN
                    SetDiagBit(6);
                    _state := E_SafeMutingState.Error;
                ELSE
                    _state := MutingStateFor(_seqIndex);
                END_IF
            ELSIF MutingEnable AND AnySensor() THEN
                // a sensor actuated out of order while muting is enabled violates the sequence
                SetDiagBit(6);
                _state := E_SafeMutingState.Error;
            ELSIF _ossdBlocked THEN
                IF Parameters.DelayTime > T#0S THEN
                    _state := E_SafeMutingState.DelayOut;
                ELSE
                    _state := E_SafeMutingState.Safe;
                END_IF
            END_IF

        E_SafeMutingState.Muting1,
        E_SafeMutingState.Muting2,
        E_SafeMutingState.Muting3,
        E_SafeMutingState.Muting4,
        E_SafeMutingState.Muting5,
        E_SafeMutingState.Muting6,
        E_SafeMutingState.Muting7,
        E_SafeMutingState.Muting8,
        E_SafeMutingState.Muting9:
            IF StateChanged() THEN
                MuteOut      := TRUE;
                MuteDelOut   := TRUE;
                MutingActive := TRUE;
            END_IF

            _maxTimer(IN := (Parameters.MaxMutingTime > T#0S), PT := Parameters.MaxMutingTime);

            IF NOT MutingEnable THEN
                // muting withdrawn: the protective device takes over immediately
                IF NOT _ossdBlocked THEN
                    _state := E_SafeMutingState.Run;
                ELSIF Parameters.DelayTime > T#0S THEN
                    _state := E_SafeMutingState.DelayOut;
                ELSE
                    _state := E_SafeMutingState.Safe;
                END_IF
            ELSIF _maxTimer.Q THEN
                SetDiagBit(7);
                _state := E_SafeMutingState.Error;
            ELSIF Advance() THEN
                SetDiagBit(6);
                _state := E_SafeMutingState.Error;
            ELSIF _seqIndex >= _seqLength THEN
                _state := E_SafeMutingState.Run;
            ELSE
                _state := MutingStateFor(_seqIndex);
            END_IF

        E_SafeMutingState.DelayOut:
            IF StateChanged() THEN
                MuteOut      := FALSE;
                MuteDelOut   := TRUE;
                MutingActive := FALSE;
                _delayTimer(IN := FALSE, PT := Parameters.DelayTime);
            END_IF

            _delayTimer(IN := TRUE, PT := Parameters.DelayTime);

            IF _delayTimer.Q THEN
                _state := SEL(_pendingError, E_SafeMutingState.Safe, E_SafeMutingState.Error);
            END_IF

        E_SafeMutingState.Error:
            IF StateChanged() THEN
                SetOutputsSafe();
                MutingActive  := FALSE;
                Error         := TRUE;
                _pendingError := FALSE;
            END_IF

            UpdateDiscrepancyDiag();

            IF _errAck AND NOT discError THEN
                _state := E_SafeMutingState.Reset;
            END_IF

        E_SafeMutingState.Reset:
            IF StateChanged() THEN
                SetOutputsSafe();
                Error := FALSE;
                Diag  := 0;
            END_IF

            IF _errAckFallingEdge THEN
                _state := SEL(_fbRun, E_SafeMutingState.Stop, E_SafeMutingState.Safe);
            END_IF
    END_CASE

    passes := passes + 1;
UNTIL (stateBefore = _state) OR (passes >= 3)
END_REPEAT

State := TO_BYTE(_state);
END_METHOD

METHOD PRIVATE SetOutputsSafe
MuteOut    := FALSE;
MuteDelOut := FALSE;
END_METHOD

METHOD PRIVATE StartEdmResetMonitoring
_edm1Dropped := FALSE;
_edm2Dropped := FALSE;
_edmResetTimer1(IN := FALSE, PT := Parameters.Edm1ResetTime);
_edmResetTimer2(IN := FALSE, PT := Parameters.Edm2ResetTime);
END_METHOD

METHOD PRIVATE StateChanged : BOOL
IF _prevState = _state THEN
    RETURN;
END_IF

_prevState   := _state;
StateChanged := TRUE;
END_METHOD

// Mirrors the discrepancy state of every pair into the diagnostic bits.
METHOD PRIVATE UpdateDiscrepancyDiag
VAR
    i : USINT;
END_VAR
FOR i := 1 TO 3 DO
    IF _pairs[i].DiscrepancyError THEN
        SetDiagBit(SEL(i = 1, SEL(i = 2, 1, 2), 0));

        IF _pairs[i].AwaitingSafeInputs THEN
            SetDiagBit(SEL(i = 1, SEL(i = 2, 9, 10), 8));
        ELSE
            ClearDiagBit(SEL(i = 1, SEL(i = 2, 9, 10), 8));
        END_IF
    END_IF
END_FOR
END_METHOD

END_FUNCTION_BLOCK

// ---- Tests/T_SafeConnection_Tests.TcPOU
FUNCTION_BLOCK T_SafeConnection_Tests EXTENDS TcUnit.FB_TestSuite
VAR
    // Test_StartsUpToDataWhenGroupRuns
    group_1 : T_SafeGroup;
    conn_1 : T_SafeConnection(group := group_1);
    i_1 : INT;
    // Test_ComErrorClearedByAcknowledge
    group_2 : T_SafeGroup;
    conn_2 : T_SafeConnection(group := group_2);
    i_2 : INT;
END_VAR

Test_StartsUpToDataWhenGroupRuns();
Test_ComErrorClearedByAcknowledge();

METHOD PRIVATE Test_ComErrorClearedByAcknowledge
VAR
    diag : BYTE;
END_VAR
TcUnit.TEST(__POUNAME());

// arrange
FOR i_2 := 1 TO 5 DO
    group_2(Run := TRUE, ErrAck := FALSE);
    conn_2(InjectComError := FALSE, StartupTime := T#0S);
END_FOR

// act
group_2(Run := TRUE, ErrAck := FALSE);
conn_2(InjectComError := TRUE, StartupTime := T#0S);
// assert
AssertEquals_BOOL(Expected := TRUE, Actual := conn_2.ComError, Message := 'com error');
AssertEquals_BOOL(Expected := FALSE, Actual := conn_2.InDataState, Message := 'dropped out of Data');
diag := conn_2.Diag AND 16#0F;
AssertEquals_BYTE(Expected := BYTE#5, Actual := diag, Message := 'diag code watchdog');
group_2(Run := TRUE, ErrAck := FALSE);
conn_2(InjectComError := FALSE, StartupTime := T#0S);
AssertEquals_BYTE(Expected := TO_BYTE(E_SafeGroupState.Error), Actual := group_2.State, Message := 'group ERROR');
group_2(Run := TRUE, ErrAck := TRUE);
conn_2(InjectComError := FALSE, StartupTime := T#0S);

FOR i_2 := 1 TO 5 DO
    group_2(Run := TRUE, ErrAck := FALSE);
    conn_2(InjectComError := FALSE, StartupTime := T#0S);
END_FOR

AssertEquals_BOOL(Expected := FALSE, Actual := conn_2.ComError, Message := 'error cleared');
AssertEquals_BOOL(Expected := TRUE, Actual := conn_2.InDataState, Message := 'restarted to Data');
TEST_FINISHED_NAMED(__POUNAME());
END_METHOD

METHOD PRIVATE Test_StartsUpToDataWhenGroupRuns
TcUnit.TEST(__POUNAME());
// act
group_1(Run := FALSE);
conn_1(StartupTime := T#0S);
AssertEquals_BOOL(Expected := TRUE, Actual := conn_1.InStartup, Message := 'in startup before the group runs');

FOR i_1 := 1 TO 5 DO
    group_1(Run := TRUE);
    conn_1(StartupTime := T#0S);
END_FOR

// assert
AssertEquals_BOOL(Expected := TRUE, Actual := conn_1.InDataState, Message := 'Data state reached');
AssertEquals_BOOL(Expected := FALSE, Actual := conn_1.InStartup, Message := 'no longer in startup');
TEST_FINISHED_NAMED(__POUNAME());
END_METHOD

END_FUNCTION_BLOCK

// ---- Tests/T_SafeInputTerminal8_Tests.TcPOU
FUNCTION_BLOCK T_SafeInputTerminal8_Tests EXTENDS TcUnit.FB_TestSuite
VAR
    // Test_SafeInputsFalseBeforeData
    group_1 : T_SafeGroup;
    terminal_1 : T_SafeInputTerminal8(group := group_1);
    // Test_SafeInputsFollowChannelsInData
    group_2 : T_SafeGroup;
    terminal_2 : T_SafeInputTerminal8(group := group_2);
    i_2 : INT;
    // Test_ComErrorForcesSafeInputsFalse
    group_3 : T_SafeGroup;
    terminal_3 : T_SafeInputTerminal8(group := group_3);
    i_3 : INT;
    // Test_RegistersAsConnection
    group_4 : T_SafeGroup;
    terminal_4 : T_SafeInputTerminal8(group := group_4);
END_VAR

Test_SafeInputsFalseBeforeData();
Test_SafeInputsFollowChannelsInData();
Test_ComErrorForcesSafeInputsFalse();
Test_RegistersAsConnection();

METHOD PRIVATE Test_SafeInputsFalseBeforeData
TcUnit.TEST(__POUNAME());

// arrange: group stopped, so the connection never reaches Data
group_1(Run := FALSE);

// act
terminal_1(Channel1 := TRUE, Channel2 := TRUE, Channel3 := TRUE, Channel4 := TRUE,
           Channel5 := TRUE, Channel6 := TRUE, Channel7 := TRUE, Channel8 := TRUE,
           StartupTime := T#0S);

// assert
AssertEquals_BOOL(Expected := FALSE, Actual := terminal_1.InDataState, Message := 'not in Data');
AssertEquals_BOOL(Expected := FALSE, Actual := terminal_1.SafeIn1, Message := 'SafeIn1 fail-safe');
AssertEquals_BOOL(Expected := FALSE, Actual := terminal_1.SafeIn2, Message := 'SafeIn2 fail-safe');
AssertEquals_BOOL(Expected := FALSE, Actual := terminal_1.SafeIn3, Message := 'SafeIn3 fail-safe');
AssertEquals_BOOL(Expected := FALSE, Actual := terminal_1.SafeIn4, Message := 'SafeIn4 fail-safe');
AssertEquals_BOOL(Expected := FALSE, Actual := terminal_1.SafeIn5, Message := 'SafeIn5 fail-safe');
AssertEquals_BOOL(Expected := FALSE, Actual := terminal_1.SafeIn6, Message := 'SafeIn6 fail-safe');
AssertEquals_BOOL(Expected := FALSE, Actual := terminal_1.SafeIn7, Message := 'SafeIn7 fail-safe');
AssertEquals_BOOL(Expected := FALSE, Actual := terminal_1.SafeIn8, Message := 'SafeIn8 fail-safe');
TEST_FINISHED_NAMED(__POUNAME());
END_METHOD

METHOD PRIVATE Test_SafeInputsFollowChannelsInData
TcUnit.TEST(__POUNAME());

// arrange: run the group until the connection is in Data
FOR i_2 := 1 TO 5 DO
    group_2(Run := TRUE);
    terminal_2(StartupTime := T#0S);
END_FOR
AssertEquals_BOOL(Expected := TRUE, Actual := terminal_2.InDataState, Message := 'Data state reached');

// act: odd channels on, even channels off
group_2(Run := TRUE);
terminal_2(Channel1 := TRUE, Channel2 := FALSE, Channel3 := TRUE, Channel4 := FALSE,
           Channel5 := TRUE, Channel6 := FALSE, Channel7 := TRUE, Channel8 := FALSE,
           StartupTime := T#0S);

// assert
AssertEquals_BOOL(Expected := TRUE, Actual := terminal_2.SafeIn1, Message := 'SafeIn1 follows Channel1');
AssertEquals_BOOL(Expected := FALSE, Actual := terminal_2.SafeIn2, Message := 'SafeIn2 follows Channel2');
AssertEquals_BOOL(Expected := TRUE, Actual := terminal_2.SafeIn3, Message := 'SafeIn3 follows Channel3');
AssertEquals_BOOL(Expected := FALSE, Actual := terminal_2.SafeIn4, Message := 'SafeIn4 follows Channel4');
AssertEquals_BOOL(Expected := TRUE, Actual := terminal_2.SafeIn5, Message := 'SafeIn5 follows Channel5');
AssertEquals_BOOL(Expected := FALSE, Actual := terminal_2.SafeIn6, Message := 'SafeIn6 follows Channel6');
AssertEquals_BOOL(Expected := TRUE, Actual := terminal_2.SafeIn7, Message := 'SafeIn7 follows Channel7');
AssertEquals_BOOL(Expected := FALSE, Actual := terminal_2.SafeIn8, Message := 'SafeIn8 follows Channel8');

// act: invert the pattern
group_2(Run := TRUE);
terminal_2(Channel1 := FALSE, Channel2 := TRUE, Channel3 := FALSE, Channel4 := TRUE,
           Channel5 := FALSE, Channel6 := TRUE, Channel7 := FALSE, Channel8 := TRUE,
           StartupTime := T#0S);

// assert
AssertEquals_BOOL(Expected := FALSE, Actual := terminal_2.SafeIn1, Message := 'SafeIn1 inverted');
AssertEquals_BOOL(Expected := TRUE, Actual := terminal_2.SafeIn2, Message := 'SafeIn2 inverted');
AssertEquals_BOOL(Expected := FALSE, Actual := terminal_2.SafeIn3, Message := 'SafeIn3 inverted');
AssertEquals_BOOL(Expected := TRUE, Actual := terminal_2.SafeIn4, Message := 'SafeIn4 inverted');
AssertEquals_BOOL(Expected := FALSE, Actual := terminal_2.SafeIn5, Message := 'SafeIn5 inverted');
AssertEquals_BOOL(Expected := TRUE, Actual := terminal_2.SafeIn6, Message := 'SafeIn6 inverted');
AssertEquals_BOOL(Expected := FALSE, Actual := terminal_2.SafeIn7, Message := 'SafeIn7 inverted');
AssertEquals_BOOL(Expected := TRUE, Actual := terminal_2.SafeIn8, Message := 'SafeIn8 inverted');
TEST_FINISHED_NAMED(__POUNAME());
END_METHOD

METHOD PRIVATE Test_ComErrorForcesSafeInputsFalse
TcUnit.TEST(__POUNAME());

// arrange: in Data with every channel on
FOR i_3 := 1 TO 5 DO
    group_3(Run := TRUE);
    terminal_3(Channel1 := TRUE, Channel2 := TRUE, Channel3 := TRUE, Channel4 := TRUE,
               Channel5 := TRUE, Channel6 := TRUE, Channel7 := TRUE, Channel8 := TRUE,
               StartupTime := T#0S);
END_FOR
AssertEquals_BOOL(Expected := TRUE, Actual := terminal_3.SafeIn8, Message := 'SafeIn8 on before the error');

// act
group_3(Run := TRUE);
terminal_3(Channel1 := TRUE, Channel2 := TRUE, Channel3 := TRUE, Channel4 := TRUE,
               Channel5 := TRUE, Channel6 := TRUE, Channel7 := TRUE, Channel8 := TRUE,
               InjectComError := TRUE, StartupTime := T#0S);

// assert
AssertEquals_BOOL(Expected := TRUE, Actual := terminal_3.ComError, Message := 'com error');
AssertEquals_BOOL(Expected := FALSE, Actual := terminal_3.SafeIn1, Message := 'SafeIn1 fail-safe on com error');
AssertEquals_BOOL(Expected := FALSE, Actual := terminal_3.SafeIn4, Message := 'SafeIn4 fail-safe on com error');
AssertEquals_BOOL(Expected := FALSE, Actual := terminal_3.SafeIn5, Message := 'SafeIn5 fail-safe on com error');
AssertEquals_BOOL(Expected := FALSE, Actual := terminal_3.SafeIn8, Message := 'SafeIn8 fail-safe on com error');
TEST_FINISHED_NAMED(__POUNAME());
END_METHOD

METHOD PRIVATE Test_RegistersAsConnection
TcUnit.TEST(__POUNAME());

// act
group_4(Run := TRUE);
terminal_4(StartupTime := T#0S);

// assert
AssertEquals_UINT(Expected := 1, Actual := group_4.ConnectionCount, Message := 'one connection registered');
AssertEquals_UINT(Expected := 0, Actual := group_4.FunctionBlockCount, Message := 'no function blocks');
TEST_FINISHED_NAMED(__POUNAME());
END_METHOD

END_FUNCTION_BLOCK

// ---- Core/T_SafeInputTerminal8.TcPOU
// Model of an eight channel safe input terminal (EL1918): a TwinSAFE connection with eight channels.
// Declare it in its group:  inputTerminal : T_SafeInputTerminal8(group := safetyGroup);
// Channel1..8 are the simulated field signals; SafeIn1..8 are what the TwinSAFE logic sees:
// forced FALSE (fail-safe) unless the connection is in the Data state.
FUNCTION_BLOCK T_SafeInputTerminal8 EXTENDS T_SafeConnection
VAR_INPUT
    Channel1 : BOOL;
    Channel2 : BOOL;
    Channel3 : BOOL;
    Channel4 : BOOL;
    Channel5 : BOOL;
    Channel6 : BOOL;
    Channel7 : BOOL;
    Channel8 : BOOL;
END_VAR
VAR_OUTPUT
    SafeIn1 : BOOL;
    SafeIn2 : BOOL;
    SafeIn3 : BOOL;
    SafeIn4 : BOOL;
    SafeIn5 : BOOL;
    SafeIn6 : BOOL;
    SafeIn7 : BOOL;
    SafeIn8 : BOOL;
END_VAR

SUPER^();
SafeIn1 := Channel1 AND InDataState;
SafeIn2 := Channel2 AND InDataState;
SafeIn3 := Channel3 AND InDataState;
SafeIn4 := Channel4 AND InDataState;
SafeIn5 := Channel5 AND InDataState;
SafeIn6 := Channel6 AND InDataState;
SafeIn7 := Channel7 AND InDataState;
SafeIn8 := Channel8 AND InDataState;

END_FUNCTION_BLOCK

// ---- Tests/T_SafeOutputTerminal2_Tests.TcPOU
FUNCTION_BLOCK T_SafeOutputTerminal2_Tests EXTENDS TcUnit.FB_TestSuite
VAR
    // Test_ChannelsFalseBeforeData
    group_1 : T_SafeGroup;
    terminal_1 : T_SafeOutputTerminal2(group := group_1);
    // Test_ChannelsFollowSafeOutsInData
    group_2 : T_SafeGroup;
    terminal_2 : T_SafeOutputTerminal2(group := group_2);
    i_2 : INT;
    // Test_ComErrorForcesChannelsFalse
    group_3 : T_SafeGroup;
    terminal_3 : T_SafeOutputTerminal2(group := group_3);
    i_3 : INT;
    // Test_RegistersAsConnection
    group_4 : T_SafeGroup;
    terminal_4 : T_SafeOutputTerminal2(group := group_4);
    // Test_GroupNotRunningForcesChannelsFalse
    group_5 : T_SafeGroup;
    terminal_5 : T_SafeOutputTerminal2(group := group_5);
    i_5 : INT;
END_VAR

Test_ChannelsFalseBeforeData();
Test_ChannelsFollowSafeOutsInData();
Test_ComErrorForcesChannelsFalse();
Test_RegistersAsConnection();
Test_GroupNotRunningForcesChannelsFalse();

METHOD PRIVATE Test_ChannelsFalseBeforeData
TcUnit.TEST(__POUNAME());

// arrange: group stopped, so the connection never reaches Data
group_1(Run := FALSE);

// act
terminal_1(SafeOut1 := TRUE, SafeOut2 := TRUE, StartupTime := T#0S);

// assert
AssertEquals_BOOL(Expected := FALSE, Actual := terminal_1.InDataState, Message := 'not in Data');
AssertEquals_BOOL(Expected := FALSE, Actual := terminal_1.Channel1, Message := 'Channel1 fail-safe');
AssertEquals_BOOL(Expected := FALSE, Actual := terminal_1.Channel2, Message := 'Channel2 fail-safe');
TEST_FINISHED_NAMED(__POUNAME());
END_METHOD

METHOD PRIVATE Test_ChannelsFollowSafeOutsInData
TcUnit.TEST(__POUNAME());

// arrange: run the group until the connection is in Data
FOR i_2 := 1 TO 5 DO
    group_2(Run := TRUE);
    terminal_2(StartupTime := T#0S);
END_FOR
AssertEquals_BOOL(Expected := TRUE, Actual := terminal_2.InDataState, Message := 'Data state reached');

// act
group_2(Run := TRUE);
terminal_2(SafeOut1 := TRUE, SafeOut2 := FALSE, StartupTime := T#0S);

